(* IEC 61131-3 sources: daoli-st-library/DL_MathData (part 7) *)

(* ---- FC_DL_WaferCountYield.st ---- *)
(*==============================================================================
 * 组件名称 (Component)  : FC_DL_WaferCountYield
 * 所属子库 (Sublibrary) : DL_MathData
 * 当前版本 (Version)    : 1.0.0
 * 兼容性 (Platform)     : CODESYS 3.5 / TwinCAT 3 / 汇川 InoProShop / Machine Expert
 *                         仅依赖纯 IEC 61131-3 标准元素，零厂商方言
 * 功能描述 (Function)   : 晶圆投入/产出/返工三计数 → 良率百分数与损失分档。
 *                         良率 = 良品/投入 x 100；分档：A 级 >= 99、B 级 >= 95、
 *                         C 级 >= 90、D 级 < 90。纯函数无状态保持。
 * 溯源 (Origin)         : 道莅 clean-room 防御性实现
 * 本文件内含 (Contains) : TYPE E_DL_YieldGrade / TYPE E_DL_WaferErr /
 *                         FUNCTION FC_DL_WaferCountYield
 * 依赖 (Depends)        : 无 DL_ 内部依赖；仅 IEC 61131-3 标准元素
 * 红线自检 (Redline)    : 无外部全局变量、无硬件地址直引 ｜ 全变量中英双语同行注释
 *                         防除零 + 无符号减法先验下界防下溢 ｜ 枚举成员全部显式赋值
 *                         纯函数无状态保持 ｜ 输出在每条早退路径前已赋确定值
 * 错误码表 (Codes)      : 16#0001_0476 故障级(否) 成功
 *                         16#0001_0477 故障级 投入计数为 0（防除零拒绝）
 *                         16#0001_0478 故障级 良品计数大于投入计数（计数矛盾）
 *                         16#0001_0479 故障级 良品+返工大于投入（计数矛盾/下溢风险）
 *                         16#0001_047A 信息级 成功但落入 D 档（不置故障标志）
 * 修订历史 (Revision)   : 2026-11-17  v1.0.0  首版入库 · R27 · 阶段三批 1
 * 验收向量 (Acceptance) : input=1000, good=995, rework=3 → 良率 99.5% → A 档 0476
 *                         input=0 → 0477；good=1001>input=1000 → 0478；
 *                         good=990+rework=20>input=1000 → 0479；input=100,good=80 → D 档 047A
 *============================================================================*)

(*-----------------------------------------------------------------------------
 * 枚举: E_DL_YieldGrade（归属 DL_MathData，损失分档结果）
 *----------------------------------------------------------------------------*)
TYPE E_DL_YieldGrade :
(
    eGradeA := 0,    // A 档：良率 >= 99% / Grade A: yield at least 99 percent
    eGradeB := 1,    // B 档：良率 >= 95% 且 < 99% / Grade B: 95 to below 99 percent
    eGradeC := 2,    // C 档：良率 >= 90% 且 < 95% / Grade C: 90 to below 95 percent
    eGradeD := 3     // D 档：良率 < 90% / Grade D: below 90 percent
);
END_TYPE

(*-----------------------------------------------------------------------------
 * 枚举: E_DL_WaferErr（归属 DL_MathData，与 FC_DL_WaferCountYield 同文件）
 *----------------------------------------------------------------------------*)
TYPE E_DL_WaferErr :
(
    eOk           := 16#0001_0476,   // 成功 / Success
    eInputZero    := 16#0001_0477,   // 故障级：投入为 0，防除零拒绝 / Fault: zero input rejected
    eGoodOverIn   := 16#0001_0478,   // 故障级：良品大于投入 / Fault: good count exceeds input
    eCountContrad := 16#0001_0479,   // 故障级：良品+返工大于投入 / Fault: good plus rework exceeds input
    eGradeDNote   := 16#0001_047A    // 信息级：成功但 D 档 / Info: success but grade D
);
END_TYPE

(*==============================================================================
 * 函数: FC_DL_WaferCountYield（纯函数，无任何状态保持）
 * 调用约定: 每周期按需调用；bValid = 计数合法且结果可用。
 *============================================================================*)
FUNCTION FC_DL_WaferCountYield : BOOL
VAR_INPUT
    uInputCnt   : UDINT;               // 投入片数 [片]，有效域 0~1.0E9 / Wafer input count [pcs]
    uOutputGood : UDINT;               // 良品片数 [片] / Good wafer count [pcs]
    uReworkCnt  : UDINT;               // 返工片数 [片] / Rework wafer count [pcs]
END_VAR
VAR_OUTPUT
    fYieldPct   : REAL;                // 良率 [百分数] / Yield [percent]
    eGrade      : E_DL_YieldGrade;     // 损失分档 A~D / Yield grade A to D
    bValid      : BOOL;                // 输入合法且结果可用标志 / Input legal and result usable flag
    eError      : E_DL_WaferErr;       // 错误码 / Error code
END_VAR
VAR CONSTANT
    DL_WFR_INPUT_MAX  : UDINT := 1000000000;  // 投入计数上限 [片] / Input count upper bound [pcs]
    DL_WFR_GRADE_A    : REAL := 99.0;         // A 档门限 [百分数] / Grade A threshold [percent]
    DL_WFR_GRADE_B    : REAL := 95.0;         // B 档门限 [百分数] / Grade B threshold [percent]
    DL_WFR_GRADE_C    : REAL := 90.0;         // C 档门限 [百分数] / Grade C threshold [percent]
    DL_WFR_PCT        : REAL := 100.0;        // 百分数系数 [百分数] / Percent factor [percent]
    DL_WFR_ZERO       : REAL := 0.0;          // 零值常量，避免裸字面量 / Zero constant
END_VAR
VAR
    fYieldCalc : REAL;                 // 良率中间量 [百分数] / Yield intermediate [percent]
    uLossCnt   : UDINT;                // 损失片数 = 投入-良品-返工（校验后计算）[片] / Loss count [pcs]
END_VAR

(*------------------------------------------------------------------------------
 * 段 1｜出口默认值：任何早退路径前输出已确定（哨兵 0 良率 + D 档 + 无效）
 *----------------------------------------------------------------------------*)
FC_DL_WaferCountYield := FALSE;                     // 返回值默认无效 / return defaults to invalid
fYieldPct := DL_WFR_ZERO;                           // 良率哨兵 0（防除零语义：保持 0）/ yield sentinel zero
eGrade := E_DL_YieldGrade.eGradeD;                  // 分档哨兵 D 档 / grade sentinel D
bValid := FALSE;                                    // 合法标志默认 FALSE / validity defaults FALSE
eError := E_DL_WaferErr.eInputZero;                 // 默认投入为 0 码 / default zero-input code

(*------------------------------------------------------------------------------
 * 段 2｜投入为 0 闸：防除零拒绝（良率保持哨兵 0）
 *----------------------------------------------------------------------------*)
IF (uInputCnt = 0) OR (uInputCnt > DL_WFR_INPUT_MAX) THEN
    eError := E_DL_WaferErr.eInputZero;             // 故障级：投入为 0 或越上限 / fault: zero or out-of-range input
    RETURN;
END_IF

(*------------------------------------------------------------------------------
 * 段 3｜计数矛盾闸：良品不得大于投入；良品+返工不得大于投入（先验下界防下溢）
 *----------------------------------------------------------------------------*)
IF uOutputGood > uInputCnt THEN
    eError := E_DL_WaferErr.eGoodOverIn;            // 故障级：良品 > 投入 / fault: good exceeds input
    RETURN;
END_IF
IF uReworkCnt > (uInputCnt - uOutputGood) THEN      // 减法前已证 input >= good，无下溢 / no underflow, proven
    eError := E_DL_WaferErr.eCountContrad;          // 故障级：良品+返工 > 投入 / fault: count contradiction
    RETURN;
END_IF

(*------------------------------------------------------------------------------
 * 段 4｜良率计算与分档：fYield = good/input x 100（除子已证非零）
 *----------------------------------------------------------------------------*)
fYieldCalc := UDINT_TO_REAL(uOutputGood) / UDINT_TO_REAL(uInputCnt) * DL_WFR_PCT;   // 良率 [百分数] / yield [percent]
IF fYieldCalc > DL_WFR_PCT THEN
    fYieldCalc := DL_WFR_PCT;                       // 上限防护（计数矛盾已拦，兜底）/ ceiling guard
END_IF
fYieldPct := fYieldCalc;                            // 输出良率 / yield output
uLossCnt := uInputCnt - uOutputGood - uReworkCnt;   // 损失片数 [片]（两条矛盾闸已保证非负）/ loss count, proven non-negative
IF fYieldPct >= DL_WFR_GRADE_A THEN
    eGrade := E_DL_YieldGrade.eGradeA;              // A 档 / grade A
    eError := E_DL_WaferErr.eOk;                    // 成功码 / success code
ELSIF fYieldPct >= DL_WFR_GRADE_B THEN
    eGrade := E_DL_YieldGrade.eGradeB;              // B 档 / grade B
    eError := E_DL_WaferErr.eOk;                    // 成功码 / success code
ELSIF fYieldPct >= DL_WFR_GRADE_C THEN
    eGrade := E_DL_YieldGrade.eGradeC;              // C 档 / grade C
    eError := E_DL_WaferErr.eOk;                    // 成功码 / success code
ELSE
    eGrade := E_DL_YieldGrade.eGradeD;              // D 档 / grade D
    eError := E_DL_WaferErr.eGradeDNote;            // 信息级：成功但 D 档（损失片数佐证）/ info: grade D note
END_IF
bValid := TRUE;                                     // 输入合法，结果可用 / input legal, result usable
FC_DL_WaferCountYield := TRUE;                      // 返回有效 / return valid
RETURN;
END_FUNCTION

(* ---- FC_DL_AbsEx.st ---- *)
(*
    FC_DL_AbsEx —— 实数绝对值防御包装（-0.0 归一、NaN/无穷拦截、极值溢出钳位）
    ------------------------------------------------------------------
    分类      : DL_MathData / Math-Exp
    前缀      : FC_DL_
    版本      : 1.0.0
    溯源      : IEC 61131-3 标准语义的道莅防御性实现
                （内部委托平台内建函数，外围统一错误码/钳位/双语文档；
                  未复制任何闭源厂商源码，参考实现仅限 MIT/Apache 许可）
    平台      : 纯 IEC 61131-3，CODESYS / TwinCAT / InoProShop 通用
    作者      : 道莅代码库 · PLC编程专家（R15）
    ------------------------------------------------------------------
    功能说明  : 求输入实数的绝对值。NaN 输入直接拦截返回 0.0 并置 16#0001_015E；
                无穷输入（超出双精度有限极值）同口径拦截归零；-0.0 归一
                为 +0.0；负数经符号取反实现，当绝对值恰为双精度极值
                1.7976931348623157E308 时按上溢口径钳位到同值并置 16#0001_022C
                （钳位值与真实绝对值一致，bValid=TRUE 降级可用）。
                全程绝不向下游输出 NaN/Inf 毒值。
    错误码    : 0000 正常 / 16#0001_015E 入参越界（NaN/无穷，已归零） / 16#0001_022C 上溢下溢（已钳位到类型极值）
    修订记录  : 2026-11-16 v1.0.0 首次入库（R15）
*)
FUNCTION FC_DL_AbsEx : LREAL
VAR_INPUT
    lrIn : LREAL; // 输入实数 [无量纲]，任意有限值或 NaN/无穷 / input real value [dimensionless], any finite value or NaN/inf
END_VAR
VAR_OUTPUT
    eErr : UDINT; // 错误码，0=正常，1=入参越界，2=上溢钳位 / error id, 0=ok, 1=input out of domain, 2=overflow clamped
    bError   : BOOL; // 是否出错，eErr 非 0 时为 TRUE / error flag, TRUE when eErr is nonzero
    bValid   : BOOL; // 输出是否有效可用，16#0001_022C 钳位降级时保持 TRUE / output valid, stays TRUE for usable clamped result of code 2
END_VAR
VAR
    lrAbs : LREAL; // 绝对值中间量 [无量纲] / intermediate absolute value [dimensionless]
END_VAR
VAR CONSTANT
    DL_AB_MAXREAL : LREAL := 1.7976931348623157E308; // 双精度有限极值 [无量纲]，超界判无穷，禁魔法数 / double precision finite max [dimensionless], beyond treated as infinity, no magic numbers
END_VAR

// 段 1｜返回值与错误状态预置，任何早退路径不留脏码 / segment 1, preset return value and error states so no early exit leaves stale codes
FC_DL_AbsEx := 0.0; // 返回值预置安全值 0.0 [无量纲] / preset return to safe value 0.0
eErr    := 16#0000_0000; // 错误码预置正常 / preset error id to ok
bError      := FALSE; // 错误标志预置无错 / preset error flag to FALSE
bValid      := TRUE; // 有效标志预置可用 / preset valid flag to TRUE

// 段 2｜非有限拦截：NaN 用自不等判据，无穷用超极值判据，一律不进取反运算 / segment 2, non-finite interception, NaN by self-inequality and infinity by bound test
IF (lrIn <> lrIn) OR (lrIn > DL_AB_MAXREAL) OR (lrIn < -DL_AB_MAXREAL) THEN
    eErr := 16#0001_015E; // 信息级：输入非有限，已归零 / informational, non-finite input, zeroed
    bError   := TRUE; // 置错误标志 / raise error flag
    bValid   := FALSE; // 输出 0.0 非真实结果，不可用 / output 0.0 is not the true result, invalid
    RETURN; // 返回预置安全值 0.0 / return preset safe value 0.0
END_IF

// 段 3｜零值归一：与 0.0 精确比较对 -0.0 与 +0.0 均成立，统一归 +0.0 / segment 3, zero normalization, exact compare catches both minus zero and plus zero
IF lrIn = 0.0 THEN
    FC_DL_AbsEx := 0.0; // -0.0 归一为 +0.0 / normalize minus zero to plus zero
    RETURN;
END_IF

// 段 4｜负数取反与极值溢出钳位 / segment 4, negation for negative input with extreme-value overflow clamp
IF lrIn < 0.0 THEN
    IF lrIn <= -DL_AB_MAXREAL THEN
        lrAbs    := DL_AB_MAXREAL; // 绝对值恰为极值，按上溢口径钳位 / magnitude at the extreme, clamped per overflow policy
        eErr := 16#0001_022C; // 上溢码：已钳位到类型极值 / overflow code, clamped to type extreme
        bError   := TRUE; // 置错误标志 / raise error flag
        // bValid 保持 TRUE：钳位值与真实绝对值一致，降级可用 / valid stays TRUE, clamped value equals the true absolute value
    ELSE
        lrAbs := -lrIn; // 域内负数直接取反 / in-domain negative input negated
    END_IF
ELSE
    lrAbs := lrIn; // 正数直通 / positive input passes through
END_IF

// 段 5｜结果非有限复检兜底（防御纵深，正常路径不可达） / segment 5, result finiteness recheck as defense in depth
IF lrAbs <> lrAbs THEN
    lrAbs    := 0.0; // 兜底安全值 / bottom-line safe value
    eErr := 16#0001_015E; // 信息级：结果异常归零 / informational, abnormal result zeroed
    bError   := TRUE; // 置错误标志 / raise error flag
    bValid   := FALSE; // 输出不可用 / output invalid
END_IF
FC_DL_AbsEx := lrAbs; // 输出绝对值 [无量纲] / output the absolute value
END_FUNCTION

(* ---- FC_DL_AcosDegChk.st ---- *)
(*==============================================================================
 * 名称 : FC_DL_AcosDegChk —— 反余弦 → 角度（输入钳位 [-1,1]，越界仍按钳位计算）
 * 分类 / 前缀 / 版本 : DL_MathData / FC_DL_ / 1.0.0
 * 溯源 : 开源语义参考（OSCAT/AixOCAT 族，MIT）或 clean-room IEC 实现，未复制源码
 * 平台 : 纯 IEC 61131-3
 * 功能说明 : 返回 acos(x) 的角度制结果 [0,180]。输入越出 [-1,1] 时钳位到
 *            边界后仍按钳位值计算（bValid=FALSE、eErr 置码提示越界），不产生
 *            NaN。恒等式 acos(x)=atan2(sqrt(1-x^2), x)（弧度）转角度输出，
 *            纯 ATAN2/SQRT 内联实现，无库内跨件依赖。
 *            边界处理：输入非有限（NaN/±Inf）置 eErr 返回 0.0（不钳位计算）。
 * 错误码 : 16#0001_1B0D = 输入越出 [-1,1]（已钳位计算），或输入非有限（NaN/±Inf）
 *          eErr=0 且 bValid=TRUE 表示输入在域内、返回值可用
 * 状态机 : R6 标注 N/A（纯函数无顺序状态，以本节替代 ELSE 兜底）
 * 红线 : R1/R2/R3 ✓ 零全局/零IO/纯IEC ｜ R4 ✓ 非有限拦截/域钳位防 NaN ｜ R10 ✓ 标准转换 ｜ R11 ✓ 分号收尾 ｜ R15 ✓ 无保留字撞名
 * 修订记录 : 2026-11-23 v1.0.0 首次入库（R76）
 *============================================================================*)
FUNCTION FC_DL_AcosDegChk : LREAL
VAR_INPUT
    fX : LREAL;    // 余弦值输入 [-1,1]，越界钳位 / cosine value input, clamped into [-1,1]
END_VAR
VAR_OUTPUT
    eErr   : UDINT;    // 故障码，0=正常，1B0D=越界钳位或非有限 / error code
    bError : BOOL;     // TRUE=本件发生故障 / TRUE when fault occurred
    bValid : BOOL;     // TRUE=输入在域内且返回值可用 / TRUE when input in domain and result usable
END_VAR
VAR
    _x  : LREAL;       // 钳位后的输入 [无量纲] / clamped input
    _fR : LREAL;       // 弧度制反余弦结果 [rad] / arccosine result in radians
END_VAR

FC_DL_AcosDegChk := 0.0;                     // 返回值预设 0.0 / preset return to zero
eErr   := 16#0000_0000;                      // 故障码清零 / clear error code
bError := FALSE;                             // 故障标志清零 / clear error flag
bValid := TRUE;                              // 预设输出可用 / preset valid flag

IF (fX <> fX) OR ((fX - fX) <> (fX - fX)) THEN    // NaN 或 ±Inf / NaN or infinite
    eErr   := 16#0001_1B0D;                  // 置非有限故障码 / set non-finite code
    bError := TRUE;                          // 置故障标志 / set error flag
    bValid := FALSE;                         // 返回值不可用 / return not usable
    RETURN;                                  // 返回 0.0 / return zero
END_IF

_x := fX;                                    // 取输入 / take input
IF _x > 1.0 THEN                             // 上越界钳位 / clamp upper
    _x := 1.0;                               // 钳到 +1 / clamp to +1
    eErr   := 16#0001_1B0D;                  // 置越界码 / set out-of-domain code
    bError := TRUE;                          // 置故障标志 / set error flag
    bValid := FALSE;                         // 提示越界（仍按钳位值出结果）/ flag clamped compute
ELSIF _x < -1.0 THEN                         // 下越界钳位 / clamp lower
    _x := -1.0;                              // 钳到 -1 / clamp to -1
    eErr   := 16#0001_1B0D;                  // 置越界码 / set out-of-domain code
    bError := TRUE;                          // 置故障标志 / set error flag
    bValid := FALSE;                         // 提示越界（仍按钳位值出结果）/ flag clamped compute
END_IF

_fR := ATAN2(SQRT(1.0 - _x * _x), _x);       // acos(x)=atan2(sqrt(1-x^2),x)，弧度 / arccosine via atan2
FC_DL_AcosDegChk := _fR * 180.0 / 3.14159265358979323846;    // 弧度转角度 / radians to degrees

END_FUNCTION

(* ---- FC_DL_AcosEx.st ---- *)
(*
    FC_DL_AcosEx —— 反余弦防御包装（定义域 [-1,1] 域闸钳位 + NaN 拦截）
    ------------------------------------------------------------------
    分类      : DL_MathData / Math-Trig
    前缀      : FC_DL_
    版本      : 1.0.0
    溯源      : IEC 61131-3 标准语义的道莅防御性实现
                （内部委托平台内建函数，外围统一错误码/钳位/双语文档；
                  未复制任何闭源厂商源码，参考实现仅限 MIT/Apache 许可）
    平台      : 纯 IEC 61131-3，CODESYS / TwinCAT / InoProShop 通用
    作者      : 道莅代码库 · PLC编程专家（R15）
    ------------------------------------------------------------------
    功能说明  : 求输入的反余弦，返回值域 [0, pi]。与 FC_DL_AsinEx 同一
                钳位策略：NaN 输入拦截返回 0.0 并置 16#0001_0172；定义域 [-1,1]
                之外（含无穷）钳位到 ±1 并置 16#0001_0172，bValid=FALSE 但仍返回
                钳位后的计算结果（0 或 pi）供降级使用；入参为 0 时结果
                pi/2 属正常域内输出不置码；域内委托内建 ACOS，结果再做
                NaN 复检兜底。
    错误码    : 0000 正常 / 16#0001_0172 入参越界（NaN 已归零，或域外已钳位到 ±1）
    修订记录  : 2026-11-16 v1.0.0 首次入库（R15）
*)
FUNCTION FC_DL_AcosEx : LREAL
VAR_INPUT
    lrIn : LREAL; // 输入实数 [无量纲]，定义域 [-1,1] / input real value [dimensionless], domain minus 1 to plus 1
END_VAR
VAR_OUTPUT
    eErr : UDINT; // 错误码，0=正常，1=入参越界（已钳位/归零） / error id, 0=ok, 1=input out of domain, clamped or zeroed
    bError   : BOOL; // 是否出错，eErr 非 0 时为 TRUE / error flag, TRUE when eErr is nonzero
    bValid   : BOOL; // 输出是否有效可用，钳位/归零降级时为 FALSE / output valid, FALSE for clamped or zeroed degraded results
END_VAR
VAR
    lrUse : LREAL; // 钳位后的实际计算入参 [无量纲] / clamped value actually fed to the kernel [dimensionless]
END_VAR
VAR CONSTANT
    DL_AC_DOM : LREAL := 1.0; // 定义域边界 [无量纲]，闭区间 / domain bound [dimensionless], closed interval
END_VAR

// 段 1｜返回值与错误状态预置，任何早退路径不留脏码 / segment 1, preset return value and error states
FC_DL_AcosEx := 0.0; // 返回值预置安全值 0.0 / preset return to safe value 0.0
eErr    := 16#0000_0000; // 错误码预置正常 / preset error id to ok
bError      := FALSE; // 错误标志预置无错 / preset error flag to FALSE
bValid      := TRUE; // 有效标志预置可用 / preset valid flag to TRUE

// 段 2｜NaN 拦截：自不等判据，归零早退，不进内核 / segment 2, NaN interception by self-inequality, zeroed early exit
IF lrIn <> lrIn THEN
    eErr := 16#0001_0172; // 信息级：输入 NaN，已归零 / informational, NaN input, zeroed
    bError   := TRUE; // 置错误标志 / raise error flag
    bValid   := FALSE; // 输出不可用 / output invalid
    RETURN; // 返回预置安全值 0.0 / return preset safe value 0.0
END_IF

// 段 3｜定义域闸门：域外（含无穷）钳位到 ±1，仍返回钳位后结果 / segment 3, domain gate, out-of-domain including infinity clamped to plus or minus 1 with result still returned
IF lrIn > DL_AC_DOM THEN
    lrUse    := DL_AC_DOM; // 上越界钳位 +1 / upper overflow clamped to plus 1
    eErr := 16#0001_0172; // 信息级：域外已钳位 / informational, out of domain clamped
    bError   := TRUE; // 置错误标志 / raise error flag
    bValid   := FALSE; // 钳位结果非真实值 / clamped result is not the true value
ELSIF lrIn < -DL_AC_DOM THEN
    lrUse    := -DL_AC_DOM; // 下越界钳位 -1 / lower overflow clamped to minus 1
    eErr := 16#0001_0172; // 信息级：域外已钳位 / informational, out of domain clamped
    bError   := TRUE; // 置错误标志 / raise error flag
    bValid   := FALSE; // 钳位结果非真实值 / clamped result is not the true value
ELSE
    lrUse := lrIn; // 域内直通（0 输入得 pi/2 属正常） / in-domain pass-through, zero input yields pi over 2 normally
END_IF

// 段 4｜委托内建 ACOS / segment 4, delegation to built-in ACOS
FC_DL_AcosEx := ACOS(lrUse); // 委托内建 ACOS 内核 / delegate to built-in ACOS kernel

// 段 5｜结果 NaN 复检兜底（防御纵深，正常路径不可达） / segment 5, result NaN recheck as defense in depth
IF FC_DL_AcosEx <> FC_DL_AcosEx THEN
    FC_DL_AcosEx := 0.0; // 兜底安全值 / bottom-line safe value
    IF eErr = 16#0000_0000 THEN
        eErr := 16#0001_0172; // 首事件优先置码 / first-event priority code
        bError   := TRUE; // 置错误标志 / raise error flag
        bValid   := FALSE; // 输出不可用 / output invalid
    END_IF
END_IF
END_FUNCTION

(* ---- FC_DL_AcosSafe.st ---- *)
(*
    FC_DL_AcosSafe —— 反余弦 Safe 族防御包装（域钳位 + bClamped 显式标志 + 委托内建）
    ------------------------------------------------------------------
    分类      : DL_MathData / Math-Trig
    前缀      : FC_DL_
    版本      : 1.0.0
    来源标签  : iec-std-wrapper（T0）
    溯源      : IEC 61131-3 标准语义的道莅防御性实现
                （内部委托平台内建 ACOS，外围钳位/错误码/双语文档；
                  未复制任何闭源厂商源码）
    平台      : 纯 IEC 61131-3，CODESYS / TwinCAT / InoProShop 通用
    分工声明  : 与 FC_DL_AsinSafe 为镜像件（ACOS 口径），与存量 FC_DL_AcosEx
                分工——AcosEx 为码位族，本件为 Safe 族样板（bClamped 显式
                钳位标志 + 16#0002 子带码位）；边界验证向量取 ±1 两点。
    作者      : 道莅代码库 · PLC 编程专家（R57）
    ------------------------------------------------------------------
    功能说明  : 求输入的反余弦，返回值域 [0, pi]。四段式防御（R45）：
                NaN 双判据拦截归零早退；|x|>1（含无穷）钳到 ±1 并置 bClamped
                仍返回钳位结果供降级（边界向量 ±1 为合法输入直通）；
                域内委托内建 ACOS；结果 NaN 复检兜底。
    错误码    : 0000 正常 / 16#0002_0001 入参非有限已归零 / 16#0002_0002 域外已钳位
    修订记录  : 2026-11-21 v1.0.0 首次入库（R57 批 2 · 序号 7）
*)
FUNCTION FC_DL_AcosSafe : LREAL
VAR_INPUT
    lrIn : LREAL; // 输入实数 [无量纲]，定义域 [-1,1] / input real value [dimensionless], domain minus one to plus one
END_VAR
VAR_OUTPUT
    eErr     : UDINT; // 错误码，0 = 正常 / error code, zero is ok
    bError   : BOOL;  // 出错标志，eErr 非 0 时为真 / error flag, true when eErr is nonzero
    bValid   : BOOL;  // 结果是否为真实值，钳位/归零降级时为假 / the result is the true value, false when degraded
    bClamped : BOOL;  // 本次调用发生定义域钳位 [-] / a domain clamp happened this call
END_VAR
VAR
    lrUse : LREAL; // 钳位后的实际计算入参 [无量纲] / the clamped value fed to the kernel [dimensionless]
END_VAR
VAR CONSTANT
    DL_ACS_DOM : LREAL := 1.0; // 定义域边界 [无量纲]，闭区间 / the domain bound [dimensionless], closed interval
END_VAR

// 段 1｜返回值与错误状态预置安全值（四段式第一段，R45）/ segment 1, preset the return and error states
FC_DL_AcosSafe := 0.0; // 返回值预置安全值 0.0 / preset the return to the safe zero
eErr     := 16#0000_0000; // 错误码预置正常 / preset the code to ok
bError   := FALSE; // 错误标志预置假 / preset the error flag false
bValid   := TRUE; // 有效标志预置真 / preset the valid flag true
bClamped := FALSE; // 钳位标志预置假 / preset the clamp flag false

// 段 2｜非有限拦截（双判据）：命中不调内建直接早退 / segment 2, the non finite interception
IF (lrIn <> lrIn) OR ((lrIn - lrIn) <> (lrIn - lrIn)) THEN // NaN 或无穷 / NaN or infinity
    eErr   := 16#0002_0001; // 信息级：输入非有限已归零 / informational, a non finite input zeroed
    bError := TRUE; // 置错误标志 / raise the error flag
    bValid := FALSE; // 输出不可用 / the output void
    RETURN; // 返回预置安全值 0.0 / return the preset safe zero
END_IF

// 段 3｜定义域闸门：域外钳到 ±1 并置 bClamped（±1 两边界点为合法输入直通）/ segment 3, the domain gate, the boundary points plus or minus one legal
IF lrIn > DL_ACS_DOM THEN // 上越界 / above the bound
    lrUse    := DL_ACS_DOM; // 钳到 +1 / clamp to plus one
    eErr     := 16#0002_0002; // 信息级：域外已钳位 / informational, clamped
    bError   := TRUE; // 置错误标志 / raise the error flag
    bValid   := FALSE; // 钳位结果非真实值 / the clamped result is not the true value
    bClamped := TRUE; // 置钳位标志 / raise the clamp flag
ELSIF lrIn < -DL_ACS_DOM THEN // 下越界 / below the bound
    lrUse    := -DL_ACS_DOM; // 钳到 -1 / clamp to minus one
    eErr     := 16#0002_0002; // 信息级：域外已钳位 / informational, clamped
    bError   := TRUE; // 置错误标志 / raise the error flag
    bValid   := FALSE; // 钳位结果非真实值 / the clamped result is not the true value
    bClamped := TRUE; // 置钳位标志 / raise the clamp flag
ELSE // 域内直通 / inside the domain
    lrUse := lrIn; // 直通 / passthrough
END_IF

// 段 4｜委托内建 ACOS（禁重实现数学内核）/ segment 4, delegation to the built-in ACOS
FC_DL_AcosSafe := ACOS(lrUse); // 委托内建内核 / delegate to the built-in kernel

// 段 5｜结果 NaN 复检兜底（防御纵深，正常路径不可达）/ segment 5, the result recheck as defense in depth
IF (FC_DL_AcosSafe <> FC_DL_AcosSafe) OR ((FC_DL_AcosSafe - FC_DL_AcosSafe) <> (FC_DL_AcosSafe - FC_DL_AcosSafe)) THEN // 结果非有限 / a non finite result
    FC_DL_AcosSafe := 0.0; // 兜底安全值 / the bottom-line safe value
    IF eErr = 16#0000_0000 THEN // 首事件优先置码 / the first event keeps the code
        eErr   := 16#0002_0001; // 信息级：结果非有限已归零 / informational, a non finite result zeroed
        bError := TRUE; // 置错误标志 / raise the error flag
        bValid := FALSE; // 输出不可用 / the output void
    END_IF
END_IF
END_FUNCTION

(* ---- FC_DL_Affine2Apply.st ---- *)
//==============================================================================
// 函数：FC_DL_Affine2Apply ｜ 中文名称：二维仿射矩阵对点坐标应用
// 所属子库：DL_MathData ｜ 版本：v1.0.0 ｜ 兼容：CODESYS V3.5+ / TwinCAT 3 / 汇川 InoProShop
// 功能描述：单片 3x3 仿射矩阵对单点坐标 (x, y) 应用变换，p' = M x [x, y, 1]^T
//           （列向量右乘，与 FC_DL_Affine2DCompose 的合成约定构成定义-应用
//           逆对：Compose 产出矩阵、Apply 消费矩阵）。现场语义：视觉像素
//           坐标到机械毫米坐标的单点映射、纠偏平台坐标换算、印刷套准偏移。
//           第三行偏差提示为本件信息级职责：喂入矩阵第三行偏离 (0, 0, 1)
//           超容差时按仿射截断（只用前两行），输出照算并提示，便于标定
//           链上游把透视矩阵误接进仿射链时尽早暴露。
// 开源溯源 (Origin)：道莅 clean-room 防御性实现（仅借 LGF 分类事实/参数域/行为定义，零代码行与符号名复制）
// 单位表：点坐标[用户单位] / 矩阵线性块[无量纲] / 平移列[用户单位]
// 错误码表：16#0001_0469 信息级（矩阵第三行偏离 (0,0,1) 超容差，按仿射截断
//           照算，不置 bError）/ 16#0001_046A 预留禁用（不得挪用）/
//           16#0001_046B 预留禁用（不得挪用）/ 16#0001_03B9 故障级（任一
//           输入非有限，或结果非有限溢出，置 bError，输出 0）/
//           16#0001_03BA 预留禁用（不得挪用）
// 状态机：N/A——纯函数无顺序状态机，无 CASE 可写，非法状态不可能出现，以头注释说明替代 ELSE 兜底
// 边界行为：① 矩阵元素或点坐标非有限（NaN 自反判 + 幅值上限兜底，R79）→
//           故障 03B9、输出 0、bValid := FALSE；② 结果非有限（大坐标乘
//           大缩放溢出）→ 复用 03B9（R90：与输入非法共用「数据不可信」
//           语义，现有输出组合不可观测出独立信息，不新占码位）；
//           ③ 第三行偏差仅提示不阻断（信息 0469），仿射截断照算；
//           ④ 失能清零不适用（纯函数无使能闸，非法输入即故障早退）；
//           ⑤ 安全侧 = 故障路径输出 0 而非原坐标，禁止未变换坐标冒充
//           已变换坐标进入下游；
//           ⑥ 恒等矩阵输入时输出等于输入（数值恒等由乘 1.0 保证，
//           非位拷贝）。
// 验收向量（算法已证，手算）：① 恒等矩阵 + (3,4) → (3,4)；② 平移
//           (10,20) + (1,1) → (11,21)；③ 旋转 90 度 + (1,0) → (0,1)。
//           编译器已证（三平台）：未跑，由收口方登记。
// 修订历史：v1.0.0 2026-11-17 首版（R24 派单 · T2-1 LGF Math 仿射变换族）
//==============================================================================

FUNCTION FC_DL_Affine2Apply : BOOL
VAR_INPUT
    afM : ARRAY[0..2, 0..2] OF LREAL;       // 仿射变换矩阵 [无量纲+用户单位混合]，行主序，p' = M x p / Affine transform matrix, row-major
    fX  : LREAL;                            // 源点 X [用户单位] / Source point X [user unit]
    fY  : LREAL;                            // 源点 Y [用户单位] / Source point Y [user unit]
END_VAR
VAR_OUTPUT
    fOutX  : LREAL;                         // 变换后 X [用户单位] / Transformed X [user unit]
    fOutY  : LREAL;                         // 变换后 Y [用户单位] / Transformed Y [user unit]
    eErr   : UDINT;                         // 错误码，0 = 无错，码位 16#0001_0469 起信息级、16#0001_03B9 起故障级（分带见错误码表） / Error code, 0 = no error, band info/fault per the code table
    bError : BOOL;                          // 故障级标志，仅故障级错误置位 / Fault-class flag, set only on fault-level codes
    bValid : BOOL;                          // 结果可用标志 / Result usable flag
END_VAR
VAR CONSTANT
    DL_A2A_EPS      : LREAL := 1.0E-6;      // 第三行偏差容差与浮点判零共用 [无量纲] / Third-row deviation and zero tolerance [dimensionless]
    DL_A2A_INF      : LREAL := 1.7976931348623157E308; // LREAL 幅值上限 / LREAL magnitude ceiling
    DL_A2A_ZERO     : LREAL := 0.0;         // 零值常量，避免裸字面量 [无量纲] / Zero constant, avoids a bare literal [dimensionless]
    DL_A2A_ONE      : LREAL := 1.0;         // 单位常量，第三行齐次项期望值 [无量纲] / Unity constant, expected homogeneous entry [dimensionless]
END_VAR
VAR
    fXt     : LREAL;                        // 第一行点积暂存 [用户单位] / First-row dot product staging
    fYt     : LREAL;                        // 第二行点积暂存 [用户单位] / Second-row dot product staging
    bNonFin : BOOL;                         // 非有限判定中间标志 / Non-finite detection intermediate flag
    nI      : INT;                          // 行循环索引 [—] / Row loop index
    nJ      : INT;                          // 列循环索引 [—] / Column loop index
END_VAR

(*------------------------------------------------------------------------------
 * 段 1｜出口默认值：返回值与输出预置（安全侧 = 0）
 *      Exit defaults: return value and outputs preset, fail-safe zero
 *-----------------------------------------------------------------------------*)
FC_DL_Affine2Apply := FALSE;                // 返回值默认无效 / Return value preset invalid
fOutX := DL_A2A_ZERO;                       // 输出 X 预置 0 / Preset X to zero
fOutY := DL_A2A_ZERO;                       // 输出 Y 预置 0 / Preset Y to zero
eErr   := 16#0000_0000;                     // 错误码先清零 / Error code cleared first
bError := FALSE;                            // 故障标志先清零 / Fault flag cleared first
bValid := FALSE;                            // 可用标志先清零 / Usable flag cleared first

(*------------------------------------------------------------------------------
 * 段 2｜输入非有限闸：矩阵九元素 + 点坐标（R79 双侧幅值判）
 *      Input non-finite gate over nine matrix entries and the point
 *-----------------------------------------------------------------------------*)
bNonFin := (fX <> fX) OR (ABS(fX) > DL_A2A_INF)
        OR (fY <> fY) OR (ABS(fY) > DL_A2A_INF); // 点坐标非有限判定 / Point non-finite check
FOR nI := 0 TO 2 DO
    FOR nJ := 0 TO 2 DO
        IF (afM[nI, nJ] <> afM[nI, nJ]) OR (ABS(afM[nI, nJ]) > DL_A2A_INF) THEN
            bNonFin := TRUE;                // 命中非有限矩阵元素 / Non-finite matrix entry hit
        END_IF
    END_FOR
END_FOR
IF bNonFin THEN
    eErr   := 16#0001_03B9;                 // 故障级：输入非有限 / Fault: non-finite input
    bError := TRUE;                         // 置故障标志（R45 配对） / Raise the fault flag
    bValid := FALSE;                        // 输出不可用 / Outputs unusable
    RETURN;                                 // 故障早退，输出保持 0 / Early return, outputs stay zero
END_IF

(*------------------------------------------------------------------------------
 * 段 3｜仿射应用：只用前两行点积（第三行截断，见段 4 提示）
 *      Affine application, first two rows only
 *-----------------------------------------------------------------------------*)
fXt := afM[0, 0] * fX + afM[0, 1] * fY + afM[0, 2]; // 第一行点积 [用户单位] / First-row dot product
fYt := afM[1, 0] * fX + afM[1, 1] * fY + afM[1, 2]; // 第二行点积 [用户单位] / Second-row dot product

(*------------------------------------------------------------------------------
 * 段 4｜第三行偏差提示：偏离 (0, 0, 1) 超容差 → 信息 0469（照算不阻断）
 *      Third-row deviation notice, computation continues
 *-----------------------------------------------------------------------------*)
IF (ABS(afM[2, 0]) > DL_A2A_EPS) OR (ABS(afM[2, 1]) > DL_A2A_EPS)
   OR (ABS(afM[2, 2] - DL_A2A_ONE) > DL_A2A_EPS) THEN
    eErr := 16#0001_0469;                   // 信息级：第三行非标准仿射，已按仿射截断 / Info: non-standard third row, affine-truncated
END_IF

(*------------------------------------------------------------------------------
 * 段 5｜结果非有限复检：大缩放乘大坐标可能溢出（复用 03B9，R90）
 *      Result non-finite recheck, code reused per R90
 *-----------------------------------------------------------------------------*)
IF (fXt <> fXt) OR (ABS(fXt) > DL_A2A_INF)
   OR (fYt <> fYt) OR (ABS(fYt) > DL_A2A_INF) THEN
    fOutX := DL_A2A_ZERO;                   // 溢出即输出 0（安全侧） / Overflow yields zero
    fOutY := DL_A2A_ZERO;                   // 溢出即输出 0 / Overflow yields zero
    eErr   := 16#0001_03B9;                 // 故障级：结果溢出复用输入非法码（R90） / Fault: overflow, code reused per R90
    bError := TRUE;                         // 置故障标志 / Raise the fault flag
    bValid := FALSE;                        // 输出不可用 / Outputs unusable
    RETURN;                                 // 故障早退 / Early return
END_IF

(*------------------------------------------------------------------------------
 * 段 6｜出口
 *      Exit
 *-----------------------------------------------------------------------------*)
fOutX := fXt;                               // 变换后 X 出口 / Transformed X outlet
fOutY := fYt;                               // 变换后 Y 出口 / Transformed Y outlet
bValid := TRUE;                             // 结果可用（含 0469 提示情形） / Result usable, including the 0469 notice case
FC_DL_Affine2Apply := TRUE;                 // 返回 TRUE = 应用有效 / Return TRUE = application valid
END_FUNCTION

(* ---- FC_DL_Affine2DChain.st ---- *)
(*
  ==================================================================
  组件名 Component  : FC_DL_Affine2DChain
  分类   Category   : DL_MathData
  复杂度 Complexity  : 中
  版本   Version    : 1.0.1
  功能   Purpose    : N 级 2D 仿射链一次合成。输入 nCount 个 3×3 齐次矩阵，按
                      固定次序合成 MOut = Mn × … × M2 × M1（列向量约定，先施加
                      M1），中间任一奇异即整体失效并置故障码，不外泄半结果。
  来源   Source     : t2-1-lgf-math（LGF Math 仿射族多级链合成）
  溯源   Origin     : 矩阵链式合成属公开线性代数语义，clean-room 自研实现（逐级
                      委托本库 FC_DL_Affine2DCompose 内核），未复制任何厂商源码。
  平台   Platform   : 纯 IEC 61131-3（仅 FOR / 数组 / 委托调用），三平台通用
  分工声明 Split     : 与 FC_DL_Affine2DCompose（两级属主）互补——后者只合成
                      两级并负责行列式相对判据；本件做 N 级链调度、退化分支与
                      链级码位装配，不重实现乘法内核、不重声明任何矩阵类型。
  依赖     Depends  : FC_DL_Affine2DCompose（DL_MathData 属主，本件逐级委托）
  作者   Author     : 道莅代码库 · PLC 编程专家（R60）
  ------------------------------------------------------------------
  边界 Boundary     :
                      一 合成次序写死列向量约定 MOut = Mn × … × M1：M1 先施加，
                         Mn 后施加；调用方若要行向量约定须自行转置，本件不设开关；
                      二 链长退化显式：nCount ≤ 0 输出单位阵并置信息级码；nCount
                         超 8 级钳位续算并置信息级码（不静默截断）；
                      三 有限性闸逐个枚举浮点输入：本件声明区 LREAL 输入集合 =
                         afMats 的 9 × nCount 个元素，闸内逐元素引用同一集合，
                         无标量 LREAL 引脚（R272 覆盖自证：9×nUsed 全枚举）；
                      四 中途奇异或中途非有限即整体失效：bValid = FALSE、输出
                         保持单位阵（不外泄半结果），故障码一次锁存于本次调用；
                      五 只读输入矩阵，不改调用方数组（PercentileLReal 纪律）。
  错误码   Codes    :
    16#0001_0620【故障级】中间阵奇异或委托内核判不可用，链合成终止
    16#0001_0621【故障级】输入矩阵含非有限元素（NaN / Inf），链合成终止
    16#0001_0622【信息级】链长越域已钳位（≤0 出单位阵，>8 钳到 8 级）
  验收   Acceptance :
    算法已证（脚本）：未跑 ｜ 编译器已证（三平台）：未跑
    V1 两级：M1 平移 (1,2)、M2 缩放 ×2 → 单位点 (0,0) 过链得 (2,4)
    V2 nCount=0 → 单位阵、bValid=TRUE、码 0622
    V3 第二级首行全零（奇异）→ bValid=FALSE、码 0620、输出仍为单位阵
  修订记录 Revision  :
    2026-11-21  v1.0.0  R60 首版（批 2 · 序号 6）
    2026-11-21  v1.0.1  R61 返修：D5 累加器改单位阵起步、逐级全委托（含
                        nUsed=1 单级链奇异判，R284）；D6 信息级 0622 两处
                        不再置 bError（R285 口径统一）
  ==================================================================
*)
FUNCTION FC_DL_Affine2DChain : BOOL
VAR_IN_OUT
    afMats : ARRAY[0..7, 0..2, 0..2] OF LREAL; // 链矩阵组 [无量纲 + 用户单位混合]，行主序，第 0 级先施加 / the chain matrices, row major, level zero applied first
END_VAR
VAR_INPUT
    nCount : DINT; // 链级数 [级]，合法域 1..8 / the chain level count, legal from one to eight
END_VAR
VAR_OUTPUT
    afMOut : ARRAY[0..2, 0..2] OF LREAL; // 合成矩阵 [无量纲 + 用户单位混合] / the composed matrix
    bValid : BOOL;                       // 结果可用标志（链中任一级失效即假）[-] / the result usable flag
    eErr   : UDINT;                      // 错误码，0 = 正常 / the error code, zero is ok
    bError : BOOL;                       // 故障锁存标志 [-] / the fault flag
END_VAR
VAR
    afAcc     : ARRAY[0..2, 0..2] OF LREAL; // 累加矩阵（当前已合成结果） / the accumulator of the composed so far
    afTmp     : ARRAY[0..2, 0..2] OF LREAL; // 本级乘积暂存（检过才接替累加器） / the staging product of this level
    afMk      : ARRAY[0..2, 0..2] OF LREAL; // 本级矩阵切片副本（三维数组不可直接切片传参） / the slice copy of this level
    nLevel    : DINT;  // 级遍历索引 [级] / the level loop index
    nI        : DINT;  // 行索引 [行] / the row index
    nJ        : DINT;  // 列索引 [列] / the column index
    nUsed     : DINT;  // 钳位后的实际级数 [级] / the clamped level count
    bAbort    : BOOL;  // 链终止标志（有限闸或奇异闸命中）[-] / the chain abort flag
    bClamped  : BOOL;  // 链长钳位标记 [-] / the level clamp flag
    bSubValid : BOOL;  // 委托内核结果可用位 [-] / the delegate usable bit
    bSubErr   : BOOL;  // 委托内核故障位 [-] / the delegate fault bit
    uSubErr   : UDINT; // 委托内核错误码 [码] / the delegate error code
END_VAR
VAR CONSTANT
    DL_A2CH_CHMAX : DINT := 8; // 链级数上界 [级]，与数组第 1 维一致 / the level bound aligned with the first dimension
END_VAR

// 段 1｜返回值与错误状态预置安全值（四段式第一段，R45）+ 输出预置单位阵 / segment 1, the preset of the return, the codes and the identity matrix
FC_DL_Affine2DChain := FALSE; // 返回值预置假 / preset the return false
bValid := FALSE; // 有效标志预置假 / preset the validity false
eErr := 16#0000_0000; // 错误码预置正常 / preset the code to ok
bError := FALSE; // 故障标志预置假 / preset the error flag false
bAbort := FALSE; // 终止标志预置假 / preset the abort flag false
bClamped := FALSE; // 钳位标记预置假 / preset the clamp flag false
bSubValid := FALSE; // 委托有效位预置假 / preset the delegate usable bit false
bSubErr := FALSE; // 委托故障位预置假 / preset the delegate fault bit false
uSubErr := 16#0000_0000; // 委托码预置零 / preset the delegate code zero
nUsed := 0; // 实际级数预置零 / preset the used level zero
FOR nI := 0 TO 2 DO // 单位阵装配 / build the identity matrix
    FOR nJ := 0 TO 2 DO // 列遍历 / the column loop
        IF nI = nJ THEN // 主对角 / the main diagonal
            afMOut[nI, nJ] := 1.0; // 对角置一 / unit on the diagonal
            afAcc[nI, nJ] := 1.0; // 累加器同步置一 / the accumulator seeded the same
        ELSE // 非对角 / the off diagonal
            afMOut[nI, nJ] := 0.0; // 非对角置零 / zero off the diagonal
            afAcc[nI, nJ] := 0.0; // 累加器同步置零 / the accumulator seeded the same
        END_IF
        afTmp[nI, nJ] := 0.0; // 暂存阵清零 / clear the staging matrix
        afMk[nI, nJ] := 0.0; // 切片副本清零 / clear the slice copy
    END_FOR
END_FOR

// 段 2｜链长域闸（退化与钳位显式，边界二）/ segment 2, the level count gate with the explicit degenerate branch
IF nCount < 1 THEN // 链长为零或负：退化为单位阵 / a non positive count degenerates to the identity
    eErr := 16#0001_0622; // 信息级：链长越域已钳位（信息级不置 bError，R285 口径统一，D6 返修）/ informational, the level count clamped, no fault bit
    bValid := TRUE; // 单位阵是合法结果 / the identity is a legal result
    FC_DL_Affine2DChain := TRUE; // 返回成功 / return success
    RETURN; // 早退：afMOut 已为单位阵（段 1 预置）/ early return with the identity already preset
END_IF
nUsed := nCount; // 域内接管级数 / take the count inside the domain
IF nUsed > DL_A2CH_CHMAX THEN // 超上界 / above the bound
    nUsed := DL_A2CH_CHMAX; // 钳到 8 级 / clamp to eight levels
    bClamped := TRUE; // 置钳位标记 / raise the clamp flag
END_IF

// 段 3｜有限性闸：9 × nUsed 个浮点元素逐个枚举（R272 覆盖自证，边界三）/ segment 3, the finiteness gate over every enumerated element
FOR nLevel := 0 TO nUsed - 1 DO // 级遍历 / the level loop
    FOR nI := 0 TO 2 DO // 行遍历 / the row loop
        FOR nJ := 0 TO 2 DO // 列遍历 / the column loop
            IF (afMats[nLevel, nI, nJ] <> afMats[nLevel, nI, nJ])
            OR ((afMats[nLevel, nI, nJ] - afMats[nLevel, nI, nJ]) <> (afMats[nLevel, nI, nJ] - afMats[nLevel, nI, nJ])) THEN // NaN 自反判 + Inf 差值自减判 / the NaN reflexive and the Inf difference tests
                bAbort := TRUE; // 置终止标志 / raise the abort flag
            END_IF
        END_FOR
    END_FOR
END_FOR
IF bAbort THEN // 输入含非有限 / a non finite input exists
    eErr := 16#0001_0621; // 故障级：输入矩阵含非有限元素 / fault grade, a non finite element in the input
    bError := TRUE; // 置错误标志（R45 配对）/ raise the error flag, paired with the fault code
    bValid := FALSE; // 结果不可用 / the result void
    RETURN; // 早退：afMOut 保持单位阵（不外泄半结果，边界四）/ early return with the identity kept
END_IF

// 段 4｜逐级合成：MOut = Mn × … × M1（累加器以单位阵起步、逐级全委托；D5 返修：nUsed=1 单级链也走一次委托补奇异判，R284）/ segment 4, the per level composition, the accumulator starts from the identity and every level is delegated
FOR nLevel := 0 TO nUsed - 1 DO // 第 0..nUsed-1 级逐级合成（单位阵为左乘起点）/ compose from level zero with the identity seeded accumulator
  IF NOT bAbort THEN // 链未终止才继续合成（终止后不再用半结果继续乘）/ compose only while the chain is alive
    afMk[0, 0] := afMats[nLevel, 0, 0]; // 切片副本第 0 行第 0 列 / slice row zero column zero
    afMk[0, 1] := afMats[nLevel, 0, 1]; // 切片副本第 0 行第 1 列 / slice row zero column one
    afMk[0, 2] := afMats[nLevel, 0, 2]; // 切片副本第 0 行第 2 列 / slice row zero column two
    afMk[1, 0] := afMats[nLevel, 1, 0]; // 切片副本第 1 行第 0 列 / slice row one column zero
    afMk[1, 1] := afMats[nLevel, 1, 1]; // 切片副本第 1 行第 1 列 / slice row one column one
    afMk[1, 2] := afMats[nLevel, 1, 2]; // 切片副本第 1 行第 2 列 / slice row one column two
    afMk[2, 0] := afMats[nLevel, 2, 0]; // 切片副本第 2 行第 0 列 / slice row two column zero
    afMk[2, 1] := afMats[nLevel, 2, 1]; // 切片副本第 2 行第 1 列 / slice row two column one
    afMk[2, 2] := afMats[nLevel, 2, 2]; // 切片副本第 2 行第 2 列 / slice row two column two
    IF NOT FC_DL_Affine2DCompose(afM1 := afAcc, afM2 := afMk, afMOut => afTmp, eErr => uSubErr, bError => bSubErr, bValid => bSubValid) THEN // 委托两级内核（含行列式相对判据；nUsed=1 时 afAcc 为单位阵，单位阵左乘精确无损，单级奇异判由本次委托补齐，D5）/ delegate the two level kernel, the identity left multiply is exact
        bAbort := TRUE; // 本级不可用 / this level is unusable
    END_IF
    IF bAbort OR (NOT bSubValid) THEN // 奇异或不可用即整体终止 / a singular or unusable level aborts the chain
        bAbort := TRUE; // 锁住终止标志 / hold the abort flag
    ELSE // 本级通过：接替累加器 / this level passed, take over the accumulator
        afAcc[0, 0] := afTmp[0, 0]; // 累加器接替第 0 行第 0 列 / take over row zero column zero
        afAcc[0, 1] := afTmp[0, 1]; // 累加器接替第 0 行第 1 列 / take over row zero column one
        afAcc[0, 2] := afTmp[0, 2]; // 累加器接替第 0 行第 2 列 / take over row zero column two
        afAcc[1, 0] := afTmp[1, 0]; // 累加器接替第 1 行第 0 列 / take over row one column zero
        afAcc[1, 1] := afTmp[1, 1]; // 累加器接替第 1 行第 1 列 / take over row one column one
        afAcc[1, 2] := afTmp[1, 2]; // 累加器接替第 1 行第 2 列 / take over row one column two
        afAcc[2, 0] := afTmp[2, 0]; // 累加器接替第 2 行第 0 列 / take over row two column zero
        afAcc[2, 1] := afTmp[2, 1]; // 累加器接替第 2 行第 1 列 / take over row two column one
        afAcc[2, 2] := afTmp[2, 2]; // 累加器接替第 2 行第 2 列 / take over row two column two
    END_IF
  END_IF
END_FOR

// 段 5｜出口装配：仅在全链通过时外泄合成阵（边界四）/ segment 5, the outlet assembly, exported only when the whole chain passed
IF bAbort THEN // 链终止 / the chain aborted
    eErr := 16#0001_0620; // 故障级：中间阵奇异或不可用 / fault grade, a singular or unusable intermediate
    bError := TRUE; // 置错误标志（R45 配对）/ raise the error flag, paired with the fault code
    bValid := FALSE; // 结果不可用 / the result void
    FC_DL_Affine2DChain := FALSE; // 返回失败（afMOut 保持单位阵）/ return failure with the identity kept
ELSE // 全链通过 / the whole chain passed
    afMOut[0, 0] := afAcc[0, 0]; // 出口第 0 行第 0 列 / outlet row zero column zero
    afMOut[0, 1] := afAcc[0, 1]; // 出口第 0 行第 1 列 / outlet row zero column one
    afMOut[0, 2] := afAcc[0, 2]; // 出口第 0 行第 2 列 / outlet row zero column two
    afMOut[1, 0] := afAcc[1, 0]; // 出口第 1 行第 0 列 / outlet row one column zero
    afMOut[1, 1] := afAcc[1, 1]; // 出口第 1 行第 1 列 / outlet row one column one
    afMOut[1, 2] := afAcc[1, 2]; // 出口第 1 行第 2 列 / outlet row one column two
    afMOut[2, 0] := afAcc[2, 0]; // 出口第 2 行第 0 列 / outlet row two column zero
    afMOut[2, 1] := afAcc[2, 1]; // 出口第 2 行第 1 列 / outlet row two column one
    afMOut[2, 2] := afAcc[2, 2]; // 出口第 2 行第 2 列 / outlet row two column two
    bValid := TRUE; // 结果可用 / the result is usable
    FC_DL_Affine2DChain := TRUE; // 返回成功 / return success
    IF bClamped THEN // 链长被钳位 / the level count was clamped
        eErr := 16#0001_0622; // 信息级：链长越域已钳位（信息级不置 bError，R285 口径统一，D6 返修）/ informational, the level count clamped, no fault bit
    END_IF
END_IF
END_FUNCTION

(* ---- FC_DL_Affine2DCompose.st ---- *)
//==============================================================================
// 函数：FC_DL_Affine2DCompose ｜ 中文名称：二维仿射变换矩阵合成
// 所属子库：DL_MathData ｜ 版本：v1.0.0 ｜ 兼容：CODESYS V3.5+ / TwinCAT 3 / 汇川 InoProShop
// 功能描述：两片 3x3 仿射矩阵按「先施加 M1、后施加 M2」的次序合成为单片
//           矩阵 MOut = M2 x M1（本库点变换约定 p' = M x p，列向量右乘），
//           单次调用内完成 3x3 乘法、行列式可逆性校验与双向非有限复检。
//           现场语义：视觉标定链的多级坐标映射（像素→机械→工件）合并为
//           单矩阵、纠偏平台级联、平移/旋转/缩放/剪切的按序合成。
//           合成次序与列向量约定为本库自有规格；行列式 |det| 小于容差判
//           不可逆，按信息级降级输出（合成结果本身仍有效，仅其逆变换
//           不可用），故障级只留给非法输入与结果溢出。
//           第三行按仿射约定忽略（不校验 0/0/1），第三行偏差提示职责
//           归 FC_DL_Affine2Apply 承担，本件不重复占用码位（R90）。
// 开源溯源 (Origin)：道莅 clean-room 防御性实现（仅借 LGF 分类事实/参数域/行为定义，零代码行与符号名复制）
// 单位表：矩阵线性块元素[无量纲]（旋转/缩放/剪切）/ 平移列元素[用户单位]
// 错误码表：16#0001_0466 信息级（合成矩阵行列式 |det| < 容差，变换不可逆，
//           结果照常输出，不置 bError）/ 16#0001_0467 预留禁用（不得挪用）/
//           16#0001_0468 预留禁用（不得挪用）/ 16#0001_03B7 故障级（任一
//           输入矩阵元素非有限，或乘积结果非有限溢出，置 bError，输出
//           零矩阵）/ 16#0001_03B8 预留禁用（不得挪用）
// 状态机：N/A——纯函数无顺序状态机，无 CASE 可写，非法状态不可能出现，以头注释说明替代 ELSE 兜底
// 边界行为：① 任一输入元素非有限（NaN 用自反判 x <> x，Inf 用幅值上限
//           兜底，R79）→ 故障 03B7、输出零矩阵、bValid := FALSE；
//           ② 乘积结果非有限（大坐标乘大缩放溢出）→ 复用 03B7（R90：
//           该场景与输入非法共用「矩阵数据不可信」语义，现有输出组合
//           不可观测出独立信息，不新占码位）、输出零矩阵；
//           ③ 行列式绝对值 < 1E-6 → 信息 0466，结果照常输出（降级
//           可观测，不置 bError）；
//           ④ 失能清零不适用（纯函数无使能闸，非法输入即故障早退）；
//           ⑤ 安全侧 = 故障路径输出零矩阵而非原矩阵，禁止半合成残阵
//           外泄到下游点应用件；
//           ⑥ 第三行不参与合成合法性判定：乘法仍按完整 3x3 执行，第三
//           行结果照算输出，调用方若喂入非标准第三行由 Apply 侧提示。
// 验收向量（算法已证，手算）：① M1=绕原点旋转 90 度、M2=平移 (10,0) →
//           MOut 平移列 = (0,10)、线性块为旋转 90 度；② M1=M2=恒等 →
//           MOut=恒等；③ M1 含缩放 (2,0.5)、M2 含剪切 k=1 → det(MOut)
//           = 2x0.5 = 1（合成保序：det(M2xM1)=det(M2)·det(M1)）。
//           编译器已证（三平台）：未跑，由收口方登记。
// 修订历史：v1.0.0 2026-11-17 首版（R24 派单 · T2-1 LGF Math 仿射变换族）
//==============================================================================

FUNCTION FC_DL_Affine2DCompose : BOOL
VAR_INPUT
    afM1 : ARRAY[0..2, 0..2] OF LREAL;      // 先施加的变换矩阵 M1 [无量纲+用户单位混合]，行主序 / First-applied transform matrix M1, row-major
    afM2 : ARRAY[0..2, 0..2] OF LREAL;      // 后施加的变换矩阵 M2 [无量纲+用户单位混合]，行主序 / Second-applied transform matrix M2, row-major
END_VAR
VAR_OUTPUT
    afMOut : ARRAY[0..2, 0..2] OF LREAL;    // 合成矩阵 MOut = M2 x M1 [无量纲+用户单位混合] / Composed matrix MOut = M2 times M1
    eErr   : UDINT;                         // 错误码，0 = 无错，码位 16#0001_0466 起信息级、16#0001_03B7 起故障级（分带见错误码表） / Error code, 0 = no error, band info/fault per the code table
    bError : BOOL;                          // 故障级标志，仅故障级错误置位 / Fault-class flag, set only on fault-level codes
    bValid : BOOL;                          // 结果可用标志 / Result usable flag
END_VAR
VAR
    afProd  : ARRAY[0..2, 0..2] OF LREAL;   // 乘积暂存阵（先算后检，检过才外泄） / Product staging array, checked before export
    nI      : INT;                          // 行循环索引 [—] / Row loop index
    nJ      : INT;                          // 列循环索引 [—] / Column loop index
    nK      : INT;                          // 求和循环索引 [—] / Summation loop index
    fAcc    : LREAL;                        // 点积累加器 [混合] / Dot-product accumulator
    fDet    : LREAL;                        // 合成矩阵线性块行列式 [无量纲] / Determinant of the composed linear block
    bNonFin : BOOL;                         // 非有限判定中间标志 / Non-finite detection intermediate flag
END_VAR
VAR CONSTANT
    DL_A2C_EPS     : LREAL := 1.0E-6;       // 行列式可逆性容差 [无量纲] / Determinant invertibility tolerance [dimensionless]
    DL_A2C_INF     : LREAL := 1.7976931348623157E308; // LREAL 幅值上限 / LREAL magnitude ceiling
    DL_A2C_ZERO    : LREAL := 0.0;          // 零值常量，避免裸字面量 [无量纲] / Zero constant, avoids a bare literal [dimensionless]
END_VAR

(*------------------------------------------------------------------------------
 * 段 1｜出口默认值：返回值与输出预置（安全侧 = 零矩阵）
 *      Exit defaults: return value and outputs preset, fail-safe zero matrix
 *-----------------------------------------------------------------------------*)
FC_DL_Affine2DCompose := FALSE;             // 返回值默认无效 / Return value preset invalid
FOR nI := 0 TO 2 DO
    FOR nJ := 0 TO 2 DO
        afMOut[nI, nJ] := DL_A2C_ZERO;      // 输出矩阵逐元素清零 / Output matrix cleared element-wise
    END_FOR
END_FOR
eErr   := 16#0000_0000;                     // 错误码先清零 / Error code cleared first
bError := FALSE;                            // 故障标志先清零 / Fault flag cleared first
bValid := FALSE;                            // 可用标志先清零 / Usable flag cleared first

(*------------------------------------------------------------------------------
 * 段 2｜输入非有限闸：两片矩阵任一元素 NaN/Inf 即拒绝（R79 双侧幅值判）
 *      Input non-finite gate over both matrices
 *-----------------------------------------------------------------------------*)
bNonFin := FALSE;                           // 非有限标志预清零 / Non-finite flag pre-cleared
FOR nI := 0 TO 2 DO
    FOR nJ := 0 TO 2 DO
        IF (afM1[nI, nJ] <> afM1[nI, nJ]) OR (ABS(afM1[nI, nJ]) > DL_A2C_INF)
           OR (afM2[nI, nJ] <> afM2[nI, nJ]) OR (ABS(afM2[nI, nJ]) > DL_A2C_INF) THEN
            bNonFin := TRUE;                // 命中非有限元素 / Non-finite element hit
        END_IF
    END_FOR
END_FOR
IF bNonFin THEN
    eErr   := 16#0001_03B7;                 // 故障级：输入矩阵元素非法 / Fault: illegal matrix element
    bError := TRUE;                         // 置故障标志（R45 配对） / Raise the fault flag
    bValid := FALSE;                        // 输出不可用 / Outputs unusable
    RETURN;                                 // 故障早退，输出保持零矩阵 / Early return, outputs stay zero
END_IF

(*------------------------------------------------------------------------------
 * 段 3｜矩阵合成：MOut = M2 x M1，完整 3x3 乘法（第三行照算不判定）
 *      Matrix composition, full 3x3 multiplication
 *-----------------------------------------------------------------------------*)
FOR nI := 0 TO 2 DO
    FOR nJ := 0 TO 2 DO
        fAcc := DL_A2C_ZERO;                // 点积累加器清零 / Accumulator cleared
        FOR nK := 0 TO 2 DO
            fAcc := fAcc + afM2[nI, nK] * afM1[nK, nJ]; // 行乘列累加 / Row-times-column accumulation
        END_FOR
        afProd[nI, nJ] := fAcc;             // 暂存乘积元素 / Stage the product element
    END_FOR
END_FOR

(*------------------------------------------------------------------------------
 * 段 4｜结果非有限复检：大坐标乘大缩放可能溢出（复用 03B7，R90）
 *      Result non-finite recheck, code reused per R90
 *-----------------------------------------------------------------------------*)
bNonFin := FALSE;                           // 非有限标志复清 / Non-finite flag re-cleared
FOR nI := 0 TO 2 DO
    FOR nJ := 0 TO 2 DO
        IF (afProd[nI, nJ] <> afProd[nI, nJ]) OR (ABS(afProd[nI, nJ]) > DL_A2C_INF) THEN
            bNonFin := TRUE;                // 命中非有限结果 / Non-finite result hit
        END_IF
    END_FOR
END_FOR
IF bNonFin THEN
    eErr   := 16#0001_03B7;                 // 故障级：结果溢出复用输入非法码（R90） / Fault: overflow, code reused per R90
    bError := TRUE;                         // 置故障标志 / Raise the fault flag
    bValid := FALSE;                        // 输出不可用 / Outputs unusable
    RETURN;                                 // 故障早退，输出保持零矩阵 / Early return, outputs stay zero
END_IF

(*------------------------------------------------------------------------------
 * 段 5｜可逆性校验：线性块行列式 |det| < 容差 → 信息级降级照常输出
 *      Invertibility check, info-level degradation with result exported
 *-----------------------------------------------------------------------------*)
fDet := afProd[0, 0] * afProd[1, 1] - afProd[0, 1] * afProd[1, 0]; // 线性块行列式 [无量纲] / Linear-block determinant
IF ABS(fDet) < DL_A2C_EPS THEN
    eErr := 16#0001_0466;                   // 信息级：合成变换不可逆（不置 bError） / Info: composed transform not invertible, no fault flag
END_IF

(*------------------------------------------------------------------------------
 * 段 6｜出口：检验通过后放行乘积阵
 *      Exit: staged product exported after checks
 *-----------------------------------------------------------------------------*)
FOR nI := 0 TO 2 DO
    FOR nJ := 0 TO 2 DO
        afMOut[nI, nJ] := afProd[nI, nJ];   // 暂存阵外泄 / Staged array exported
    END_FOR
END_FOR
bValid := TRUE;                             // 结果可用（含 0466 降级情形） / Result usable, including the degraded case
FC_DL_Affine2DCompose := TRUE;              // 返回 TRUE = 合成有效 / Return TRUE = composition valid
END_FUNCTION

(* ---- FC_DL_Affine2DInvert.st ---- *)
//==============================================================================
// 函数：FC_DL_Affine2DInvert ｜ 中文名称：二维仿射变换矩阵求逆
// 所属子库：DL_MathData ｜ 版本：v1.0.0 ｜ 兼容：CODESYS V3.5+ / TwinCAT 3 / 汇川 InoProShop
// 功能描述：3x3 仿射矩阵求逆——线性块取 2x2 伴随/行列式法，平移列按
//           t' = -A^(-1) x t 反算；点变换约定沿用本库 p' = M x p（列向量
//           右乘、行主序存储）。与 FC_DL_Affine2DCompose / FC_DL_Affine2DApply
//           构成定义-应用-逆三元闭环。与 Compose 的「不可逆降级照算」策略
//           分立：本件不可逆时输出全零矩阵，禁止半逆残阵外泄（半逆会被
//           下游点应用件当成有效映射，标定链错位难查）。库内已有
//           FC_DL_Matrix3Inverse，但其行列式含第三行，与仿射语义（第三行
//           恒为 0/0/1）不等价，按「库内委托须等价」纪律不委托、就地实现。
// 开源溯源 (Origin)：道莅 clean-room 防御性实现（仅借 LGF 分类事实/参数域/行为定义，零代码行与符号名复制）
// 单位表：矩阵线性块元素[无量纲]（旋转/缩放/剪切）/ 平移列元素[用户单位] / 行列式[无量纲]
// 错误码表：16#0001_046F 信息级（线性块奇异 |det| 小于相对判据，不可逆，
//           输出全零矩阵，不置 bError）/ 16#0001_0470 预留禁用（不得挪用）/
//           16#0001_03BD 故障级（任一输入元素非有限，或求逆结果非有限
//           溢出，置 bError，输出全零矩阵）/ 16#0001_03BE 预留禁用（不得挪用）
// 状态机：N/A——纯函数无顺序状态机，无 CASE 可写，非法状态不可能出现，以头注释说明替代 ELSE 兜底
// 边界行为：① 任一输入元素非有限（NaN 用自反判 x <> x，Inf 用幅值上限
//           兜底，R79）→ 故障 03BD、afMInv 全 0、bValid := FALSE；
//           ② |det| 小于等于 fDetEps 乘线性块最大绝对值平方（相对判据，
//           R13 Matrix3Inverse 口径）→ 信息 046F、afMInv 全 0、bValid :=
//           FALSE——不可逆禁止半逆外泄，与 Compose 降级照算策略分立；
//           ③ 第三行不参与求逆（R90 家族）：行列式与逆只按 2x2 线性块
//           加平移列计算，输出第三行按输入第三行原样回填，不做 0/0/1
//           校验（偏差提示职责归 Apply 侧，本件不重复占码位）；
//           ④ fDetEps 非正 → 回退默认 1.0E-6（容差引脚自愈，不置错）；
//           ⑤ 求逆结果非有限（大坐标乘大缩放溢出）→ 复用 03BD（R90：
//           与输入非法共用「矩阵数据不可信」语义，现有输出组合不可观测
//           出独立信息，不新占码位）、afMInv 全 0；
//           ⑥ 安全侧 = 故障与不可逆路径输出全零矩阵而非原矩阵或残阵；
//           ⑦ 失能清零不适用（纯函数无使能闸，非法输入即故障早退）。
// 修订历史：v1.0.0 2026-11-17 首版（R25 派单 · §4.1）
//==============================================================================
FUNCTION FC_DL_Affine2DInvert : BOOL
VAR_INPUT
    afM     : ARRAY[0..2, 0..2] OF LREAL;   // 待求逆仿射矩阵 M [无量纲+用户单位混合]，行主序 / Affine matrix M to invert, row-major
    fDetEps : LREAL := 1.0E-6;              // 相对奇异判据 [无量纲]，非正回退默认 / Relative singularity threshold, non-positive falls back to default
END_VAR
VAR_OUTPUT
    afMInv  : ARRAY[0..2, 0..2] OF LREAL;   // 逆矩阵 M^(-1) [无量纲+用户单位混合]，失败时全 0 / Inverse matrix, all zero on failure
    fDet    : LREAL;                        // 线性块行列式 [无量纲] / Determinant of the linear block
    eErr    : UDINT;                        // 错误码，0 = 无错，码位 16#0001_046F 起信息级、16#0001_03BD 起故障级（分带见错误码表） / Error code, 0 = no error, band info/fault per the code table
    bError  : BOOL;                         // 故障级标志，仅故障级错误置位 / Fault-class flag, set only on fault-level codes
    bValid  : BOOL;                         // 结果可用标志，不可逆与非有限路径显式 FALSE / Result usable flag, explicit FALSE on singular and non-finite paths
END_VAR
VAR
    nI      : INT;                          // 行循环索引 [—] / Row loop index
    nJ      : INT;                          // 列循环索引 [—] / Column loop index
    fMaxAbs : LREAL;                        // 线性块元素绝对值最大值 [无量纲] / Max absolute value of the linear block
    fAbsK   : LREAL;                        // 当前元素绝对值暂存 [无量纲] / Absolute value of the current element
    fEpsEff : LREAL;                        // 生效奇异判据 [无量纲] / Effective singularity threshold
    fInv00  : LREAL;                        // 逆线性块 (0,0) 元素暂存 [无量纲] / Inverse linear block element (0,0)
    fInv01  : LREAL;                        // 逆线性块 (0,1) 元素暂存 [无量纲] / Inverse linear block element (0,1)
    fInv10  : LREAL;                        // 逆线性块 (1,0) 元素暂存 [无量纲] / Inverse linear block element (1,0)
    fInv11  : LREAL;                        // 逆线性块 (1,1) 元素暂存 [无量纲] / Inverse linear block element (1,1)
    fInv02  : LREAL;                        // 逆平移列 x 分量暂存 [用户单位] / Inverse translation x component
    fInv12  : LREAL;                        // 逆平移列 y 分量暂存 [用户单位] / Inverse translation y component
    bNonFin : BOOL;                         // 非有限判定中间标志 / Non-finite detection intermediate flag
END_VAR
VAR CONSTANT
    DL_A2I_CODE_INFO_1 : UDINT := 16#0001_046F;   // 信息级槽 1（线性块奇异） / info slot 1
    DL_A2I_CODE_INFO_2 : UDINT := 16#0001_0470;   // 预留禁用（不得挪用） / reserved, do not use
    DL_A2I_CODE_FLT_1  : UDINT := 16#0001_03BD;   // 故障级槽 1（输入元素非有限） / fault slot 1
    DL_A2I_CODE_FLT_2  : UDINT := 16#0001_03BE;   // 预留禁用（不得挪用） / reserved, do not use
    DL_A2I_EPS_DEF : LREAL := 1.0E-6;               // 默认相对奇异判据 [无量纲] / Default relative singularity threshold [dimensionless]
    DL_A2I_INF     : LREAL := 1.7976931348623157E308; // LREAL 幅值上限，Inf 判据 / LREAL magnitude ceiling, Inf criterion
    DL_A2I_ZERO    : LREAL := 0.0;                  // 零值常量，避免裸字面量 [无量纲] / Zero constant, avoids a bare literal [dimensionless]
END_VAR

(*------------------------------------------------------------------------------
 * 段 1｜出口默认值先行：全零矩阵 + 无错 + 不可用（先写后算，任何早退路径出口确定）
 *----------------------------------------------------------------------------*)
FOR nI := 0 TO 2 DO
    FOR nJ := 0 TO 2 DO
        afMInv[nI, nJ] := DL_A2I_ZERO;         // 逆矩阵默认全零 / default all-zero inverse
    END_FOR
END_FOR
fDet   := DL_A2I_ZERO;                         // 行列式默认零 / determinant defaults to zero
eErr   := 16#0000_0000;                        // 错误码默认无错 / error code defaults to none
bError := FALSE;                               // 故障标志默认清除 / fault flag cleared
bValid := FALSE;                               // 可用标志默认不可用，算完并检过才置位 / usable flag FALSE until computed and checked

(*------------------------------------------------------------------------------
 * 段 2｜输入非有限全阵扫描（9 元素逐个：NaN 自反判 + Inf 幅值上限判，R79）
 *----------------------------------------------------------------------------*)
bNonFin := FALSE;                              // 非有限标志复位 / reset non-finite flag
FOR nI := 0 TO 2 DO
    FOR nJ := 0 TO 2 DO
        IF (afM[nI, nJ] <> afM[nI, nJ]) OR (ABS(afM[nI, nJ]) >= DL_A2I_INF) THEN
            bNonFin := TRUE;                   // 发现非有限元素 / non-finite element found
        END_IF
    END_FOR
END_FOR
IF bNonFin THEN
    eErr   := DL_A2I_CODE_FLT_1;               // 故障级：任一输入元素非有限 / fault: non-finite input element
    bError := TRUE;                            // 故障级必置 bError（R45 配对）/ fault-class pairs with bError
    bValid := FALSE;                           // 输出不可用 / outputs unusable
    FC_DL_Affine2DInvert := FALSE;             // 返回值 = 可用标志同口径 / return mirrors bValid
    RETURN;
END_IF

(*------------------------------------------------------------------------------
 * 段 3｜线性块行列式与相对奇异判据（第三行不参与，R90 家族）
 *----------------------------------------------------------------------------*)
fDet := afM[0, 0] * afM[1, 1] - afM[0, 1] * afM[1, 0];  // 2x2 线性块行列式 / 2x2 linear block determinant
fMaxAbs := ABS(afM[0, 0]);                     // 最大绝对值种子：m00 / seed max with m00
fAbsK := ABS(afM[0, 1]);                       // m01 绝对值 / absolute of m01
IF fAbsK > fMaxAbs THEN fMaxAbs := fAbsK; END_IF
fAbsK := ABS(afM[1, 0]);                       // m10 绝对值 / absolute of m10
IF fAbsK > fMaxAbs THEN fMaxAbs := fAbsK; END_IF
fAbsK := ABS(afM[1, 1]);                       // m11 绝对值 / absolute of m11
IF fAbsK > fMaxAbs THEN fMaxAbs := fAbsK; END_IF
fEpsEff := fDetEps;                            // 生效判据先取引脚 / effective threshold from pin
IF fEpsEff <= DL_A2I_ZERO THEN
    fEpsEff := DL_A2I_EPS_DEF;                 // 非正回退默认判据 / non-positive falls back to default
END_IF
IF ABS(fDet) <= fEpsEff * fMaxAbs * fMaxAbs THEN
    eErr   := DL_A2I_CODE_INFO_1;              // 信息级：线性块奇异，不可逆 / info: singular linear block, not invertible
    bError := FALSE;                           // 信息级不置 bError（R45/R101）/ info never raises bError
    bValid := FALSE;                           // 逆矩阵不可用，禁止半逆外泄 / inverse unusable, no half-inverse leak
    FC_DL_Affine2DInvert := FALSE;             // 返回值同口径 / return mirrors bValid
    RETURN;
END_IF

(*------------------------------------------------------------------------------
 * 段 4｜2x2 伴随求逆 + 平移列反算 t' = -A^(-1) x t（除子 fDet 已由段 3 保证非零）
 *----------------------------------------------------------------------------*)
fInv00 :=  afM[1, 1] / fDet;                   // A^(-1)(0,0) = m11/det / inverse element
fInv01 := -afM[0, 1] / fDet;                   // A^(-1)(0,1) = -m01/det / inverse element
fInv10 := -afM[1, 0] / fDet;                   // A^(-1)(1,0) = -m10/det / inverse element
fInv11 :=  afM[0, 0] / fDet;                   // A^(-1)(1,1) = m00/det / inverse element
fInv02 := -(fInv00 * afM[0, 2] + fInv01 * afM[1, 2]);  // 逆平移列 x = -(A^(-1) x t)_x / inverse translation x
fInv12 := -(fInv10 * afM[0, 2] + fInv11 * afM[1, 2]);  // 逆平移列 y = -(A^(-1) x t)_y / inverse translation y

(*------------------------------------------------------------------------------
 * 段 5｜结果非有限复检（溢出复用 03BD，见边界行为⑤）后装配输出
 *----------------------------------------------------------------------------*)
IF (fInv00 <> fInv00) OR (fInv01 <> fInv01) OR (fInv10 <> fInv10) OR (fInv11 <> fInv11)
   OR (fInv02 <> fInv02) OR (fInv12 <> fInv12)
   OR (ABS(fInv00) >= DL_A2I_INF) OR (ABS(fInv01) >= DL_A2I_INF)
   OR (ABS(fInv10) >= DL_A2I_INF) OR (ABS(fInv11) >= DL_A2I_INF)
   OR (ABS(fInv02) >= DL_A2I_INF) OR (ABS(fInv12) >= DL_A2I_INF) THEN
    FOR nI := 0 TO 2 DO
        FOR nJ := 0 TO 2 DO
            afMInv[nI, nJ] := DL_A2I_ZERO;     // 溢出路径安全侧：全零矩阵 / overflow path safe side: all-zero
        END_FOR
    END_FOR
    eErr   := DL_A2I_CODE_FLT_1;               // 故障级：求逆结果非有限溢出 / fault: non-finite inverse result
    bError := TRUE;                            // 故障级必置 bError（R45 配对）/ fault-class pairs with bError
    bValid := FALSE;                           // 输出不可用 / outputs unusable
    FC_DL_Affine2DInvert := FALSE;             // 返回值同口径 / return mirrors bValid
    RETURN;
END_IF

(*------------------------------------------------------------------------------
 * 段 6｜装配输出：线性块 + 平移列 + 第三行原样回填（边界行为③）
 *----------------------------------------------------------------------------*)
afMInv[0, 0] := fInv00;                        // 逆线性块 (0,0) / inverse element
afMInv[0, 1] := fInv01;                        // 逆线性块 (0,1) / inverse element
afMInv[0, 2] := fInv02;                        // 逆平移列 x / inverse translation x
afMInv[1, 0] := fInv10;                        // 逆线性块 (1,0) / inverse element
afMInv[1, 1] := fInv11;                        // 逆线性块 (1,1) / inverse element
afMInv[1, 2] := fInv12;                        // 逆平移列 y / inverse translation y
afMInv[2, 0] := afM[2, 0];                     // 第三行原样回填，不校验 / third row copied verbatim, unchecked
afMInv[2, 1] := afM[2, 1];                     // 第三行原样回填，不校验 / third row copied verbatim, unchecked
afMInv[2, 2] := afM[2, 2];                     // 第三行原样回填，不校验 / third row copied verbatim, unchecked
eErr   := 16#0000_0000;                        // 无错出口 / no-error exit
bError := FALSE;                               // 无故障 / no fault
bValid := TRUE;                                // 逆矩阵可用 / inverse usable
FC_DL_Affine2DInvert := TRUE;                  // 返回值 = 可用标志 / return mirrors bValid
END_FUNCTION

(* ---- FC_DL_AffineTransformPoint.st ---- *)
(*
    FC_DL_AffineTransformPoint —— 2D 仿射点变换
    ------------------------------------------------------------------
    分类      : DL_MathData / Transform
    前缀      : FC_DL_
    版本      : 1.0.0
    溯源      : T2-1 LGF · Math（源矩阵明列「仿射变换组合族待挖」；只借该族归属
                Math 的分类事实）；旋转 / 缩放 / 平移的合成顺序为本库自有规格，
                角度归一式的工程写法、码位与错误分级 100% 自有；
                clean-room 重写，未复制任何闭源厂商源码，参考实现仅限 MIT/Apache 许可
    平台      : 纯 IEC 61131-3，CODESYS V3.5+ / TwinCAT 3 / InoProShop 通用
    作者      : 道莅代码库 · PLC编程专家（R18）
    ------------------------------------------------------------------
    功能说明  : 单次完成「绕原点旋转 → 各轴缩放 → 平移」的合成，输出变换后坐标。
                现场语义：视觉像素坐标到机械 mm 坐标（含相机安装角偏差）、纠偏平台
                坐标映射、印刷套准偏移换算；
                角度归一用「减 360 乘整数商」单算式路径，不用循环也不用取余
                （浮点取余在三平台行为不一致）；三角函数直接调用内建 SIN / COS，
                绝不重实现（T0 判据 2）；
                缩放为 0 使变换不可逆，按故障拒绝并原值回送，绝不返回被压平的点；
                输入与中间结果双向非有限复检，1e38 量级缩放乘大坐标的溢出能被抓住。
    错误码    : 16#0001_0241 旋转角超正负 360 度已归一——信息级，正常防御
                16#0001_0242 预留禁用（信息级，不得挪用）
                16#0001_0318 缩放因子为 0（变换不可逆）——故障级，返回原点值
                16#0001_0319 输入或中间结果非有限（NaN / 正负 INF / 溢出）——故障级，输出 0
                16#0001_031A 预留禁用（故障级，不得挪用）
    码位总账  : 16#0001_0241 用 / 16#0001_0242 预留 ｜ 16#0001_0318 用 / 16#0001_0319 用 / 16#0001_031A 预留
    状态机    : N/A —— 纯函数无顺序状态机，无 CASE 可写，非法状态不可能出现
    采样约定  : 纯组合函数，无定时器、无内部驻留状态；变换参数由调用方保证在同一
                标定批次内恒定（本库统一约定：标定参数只在停机态下发）。
    修订记录  : 2026-11-16 v1.0.0 首次入库（R18）
*)
FUNCTION FC_DL_AffineTransformPoint : BOOL
VAR_INPUT
    fX       : REAL := 0.0;                    // 源点 X [用户单位] / source point X [user unit]
    fY       : REAL := 0.0;                    // 源点 Y [用户单位] / source point Y [user unit]
    fRotDeg  : REAL := 0.0;                    // 旋转角，正为逆时针 [度]，范围 -720.0~720.0 / rotation angle, positive counter clockwise [deg], range -720.0~720.0
    fScaleX  : REAL := 1.0;                    // X 缩放比 [比值]，范围 0.001~1000.0，禁 0 / X scale ratio [ratio], range 0.001~1000.0, zero forbidden
    fScaleY  : REAL := 1.0;                    // Y 缩放比 [比值]，范围 0.001~1000.0，禁 0 / Y scale ratio [ratio], range 0.001~1000.0, zero forbidden
    fTx      : REAL := 0.0;                    // X 平移量 [用户单位] / X translation [user unit]
    fTy      : REAL := 0.0;                    // Y 平移量 [用户单位] / Y translation [user unit]
END_VAR
VAR_OUTPUT
    fOutX  : REAL;                             // 变换后 X [用户单位] / transformed X [user unit]
    fOutY  : REAL;                             // 变换后 Y [用户单位] / transformed Y [user unit]
    eErr   : UDINT;                            // 错误码，0=正常 / error id, 0=ok
    bError : BOOL;                             // 故障标志，eErr 为故障级时 TRUE / error flag, TRUE on fault-level eErr
    bValid : BOOL;                             // 结果是否可用 / result usable flag
END_VAR
VAR
    fAngNorm : REAL;                           // 归一后角度 [度]，范围 0~360 / normalised angle [deg], range 0~360
    fRad     : REAL;                           // 归一后角度换算的弧度 [弧度] / normalised angle in radians [rad]
    fCos     : REAL;                           // 余弦值，范围 -1.0~1.0 [无量纲] / cosine value, range -1.0~1.0 [dimensionless]
    fSin     : REAL;                           // 正弦值，范围 -1.0~1.0 [无量纲] / sine value, range -1.0~1.0 [dimensionless]
    fXRot    : REAL;                           // 旋转后 X [用户单位] / X after rotation [user unit]
    fYRot    : REAL;                           // 旋转后 Y [用户单位] / Y after rotation [user unit]
    fXScaled : REAL;                           // 缩放后 X [用户单位] / X after scaling [user unit]
    fYScaled : REAL;                           // 缩放后 Y [用户单位] / Y after scaling [user unit]
    fQuot    : REAL;                           // 角度除以 360 的整数商中间量 [无量纲] / integer quotient of the angle divided by 360 [dimensionless]
    bNonFin  : BOOL;                           // 非有限判定中间标志 / non-finite detection intermediate flag
END_VAR
VAR CONSTANT
    DL_AFF_EPS        : REAL := 1.0E-6;        // 浮点判等容差 [无量纲] / float equality tolerance [dimensionless]
    DL_AFF_INF_GUARD  : REAL := 4.0E38;        // 非有限幅值判定阈值，高于 REAL 最大有限值 [用户单位] / non-finite magnitude guard above the largest finite REAL [user unit]
    DL_AFF_FULL_DEG   : REAL := 360.0;         // 一整圈角度 [度] / one full turn [deg]
    DL_AFF_DEG2RAD    : REAL := 0.017453292519943295; // 度转弧度系数 [弧度每度] / degree to radian factor [rad per deg]
    DL_AFF_ZERO       : REAL := 0.0;           // 零值常量，避免裸字面量 [无量纲] / zero constant, avoids a bare literal [dimensionless]
    DL_AFF_TWO        : REAL := 2.0;           // 除数二，用于半圆判定 [无量纲] / divisor two, used by the half turn check [dimensionless]
END_VAR

// 段 1｜返回值与输出预置 / segment 1, preset return value and outputs
FC_DL_AffineTransformPoint := FALSE;           // 故障缺省返回 FALSE / fault default returns FALSE
fOutX := DL_AFF_ZERO;                          // 输出 X 预置 0 / preset X to zero
fOutY := DL_AFF_ZERO;                          // 输出 Y 预置 0 / preset Y to zero
eErr := 0;                                     // 预置无错误 / preset no error
bError := FALSE;                               // 预置无故障 / preset no fault
bValid := FALSE;                               // 预置结果不可用 / preset unusable

// 段 2｜输入非有限闸：任一输入 NaN 或正负 INF 即拒绝 / segment 2, input non-finite gate
bNonFin := (fX <> fX) OR (fX > DL_AFF_INF_GUARD) OR (fX < -DL_AFF_INF_GUARD)
        OR (fY <> fY) OR (fY > DL_AFF_INF_GUARD) OR (fY < -DL_AFF_INF_GUARD)
        OR (fRotDeg <> fRotDeg) OR (fRotDeg > DL_AFF_INF_GUARD) OR (fRotDeg < -DL_AFF_INF_GUARD)
        OR (fTx <> fTx) OR (fTx > DL_AFF_INF_GUARD) OR (fTx < -DL_AFF_INF_GUARD)
        OR (fTy <> fTy) OR (fTy > DL_AFF_INF_GUARD) OR (fTy < -DL_AFF_INF_GUARD); // 平移与角度同样检查 / translation and angle are checked the same way
IF bNonFin THEN
    eErr := 16#0001_0319;                      // 输入非有限故障码 / non-finite input fault id
    bError := TRUE;                            // 置故障标志 / raise the error flag
    RETURN;                                    // 故障级提前返回，输出保持 0 / early return on fault, outputs stay zero
END_IF

// 段 3｜缩放闸：缩放为 0 使变换不可逆，原值回送并拒绝 / segment 3, zero scale gate
IF (ABS(fScaleX) < DL_AFF_EPS) OR (ABS(fScaleY) < DL_AFF_EPS) THEN
    eErr := 16#0001_0318;                      // 缩放为零故障码 / zero scale fault id
    bError := TRUE;                            // 置故障标志 / raise the error flag
    fOutX := fX;                               // 原值回送 X，便于上层诊断 / return the original X so the caller can diagnose
    fOutY := fY;                               // 原值回送 Y / return the original Y
    RETURN;                                    // 故障级提前返回 / early return on fault
END_IF

// 段 4｜角度归一：减 360 乘以整数商，单算式路径，不用循环也不用取余 / segment 4, angle normalisation
fAngNorm := fRotDeg;                           // 默认沿用输入角 / default to the input angle
IF ABS(fRotDeg) > DL_AFF_FULL_DEG THEN
    fQuot := TRUNC(fRotDeg / DL_AFF_FULL_DEG); // 整数商（向零截断，除数为常量 360 恒非零）/ integer quotient, truncated toward zero, the divisor is the constant 360
    fAngNorm := fRotDeg - DL_AFF_FULL_DEG * fQuot; // 单算式归一，残差落在正负 360 内 / single expression normalisation, the residual stays within plus or minus 360
    eErr := 16#0001_0241;                      // 归一提示（信息级不置故障）/ normalisation hint, info level never raises a fault
END_IF

// 段 5｜三角函数：直接调内建，绝不重实现 / segment 5, trigonometric functions are built-in calls only
fRad := fAngNorm * DL_AFF_DEG2RAD;             // 度转弧度 / degrees to radians
fCos := COS(fRad);                             // 余弦 [无量纲] / cosine [dimensionless]
fSin := SIN(fRad);                             // 正弦 [无量纲] / sine [dimensionless]

// 段 6｜旋转 → 缩放 → 平移 合成 / segment 6, rotation then scaling then translation
fXRot := fX * fCos - fY * fSin;                // 旋转后 X / X after rotation
fYRot := fX * fSin + fY * fCos;                // 旋转后 Y / Y after rotation
fXScaled := fXRot * fScaleX;                   // 各轴缩放 X / per axis scaling on X
fYScaled := fYRot * fScaleY;                   // 各轴缩放 Y / per axis scaling on Y
fOutX := fXScaled + fTx;                       // 叠加 X 平移 / add the X translation
fOutY := fYScaled + fTy;                       // 叠加 Y 平移 / add the Y translation

// 段 7｜结果非有限复检：大缩放乘大坐标可能溢出 / segment 7, result non-finite recheck
bNonFin := (fOutX <> fOutX) OR (fOutX > DL_AFF_INF_GUARD) OR (fOutX < -DL_AFF_INF_GUARD)
        OR (fOutY <> fOutY) OR (fOutY > DL_AFF_INF_GUARD) OR (fOutY < -DL_AFF_INF_GUARD); // 结果溢出判定 / result overflow check
IF bNonFin THEN
    fOutX := DL_AFF_ZERO;                      // 溢出即输出 0 / overflow yields zero
    fOutY := DL_AFF_ZERO;                      // 溢出即输出 0 / overflow yields zero
    eErr := 16#0001_0319;                      // 结果非有限故障码 / non-finite result fault id
    bError := TRUE;                            // 置故障标志 / raise the error flag
    RETURN;                                    // 故障级提前返回 / early return on fault
END_IF

// 段 8｜出口 / segment 8, exit
bValid := TRUE;                                // 结果可用 / the result is usable
FC_DL_AffineTransformPoint := TRUE;            // 变换成功 / the transform succeeded
END_FUNCTION

(* ---- FC_DL_AkimaInterp1D.st ---- *)
(*
  道莅工业代码库 | DL_MathData | FC_DL_AkimaInterp1D
  版本: 1.0.0 | 日期: 2026-11-23 | 轮次: R75
  开源溯源: self-cleanroom（无外部来源；Akima 1970 抗振荡插值为公开算法，
            本件独立实现，零代码行复制）
  功能: Akima 一维插值（显式点数入参防 VLA）——5 点及以上走完整 Akima
        切线加权（端部斜率外推两支），2~4 点回落线性插值；查询点越界钳端点。
  兼容性: CODESYS 3.5 / TwinCAT 3 / 汇川 InoProShop；仅依赖标准 ABS/SQRT，零厂商私有库
  接口: 输入查询点 fX、节点表 aX/aY（固定上界 ARRAY[1..100] OF REAL）、
        uPointCnt（1..200，内部钳位 [2,100]）；返回值 TRUE=已执行；
        输出 fY（越界钳端点值）、bValid、eErr。纯函数：无内部状态。
  码表: 16#0001_0500 故障级：节点表非法（含非有限值或未严格升序，或查询点 NaN）
        码段说明：0001 段 03xx 故障子带已满（03FF 已占用），启用 05xx 扩展域闸子带，
        0500 槽经全库实扫空闲。
  边界: ① uPointCnt 先钳位 [2,100]（R75 显式点数字段口径），钳位后 < 2 不可能，
        表非法仅由升序破坏/非有限/查询 NaN 触发；
        ② 段斜率除法分母由升序闸（节点差 > EPS）证明 > 0；
        ③ Akima 切线权重分母 (w1+w2) = 0 时回落两邻段斜率均值（算法标准防除零）；
        ④ 端部外推斜率 m0/m-1/mn/mn+1 需 n >= 4，本件以 n >= 5 进 Akima 路径闸住；
        ⑤ 全部输出在所有路径（含提前返回）赋值；⑥ 零全局耦合。
  邻件比对: Lagrange/Hermite/CubicSpline（多项式样条族 vs 本件 Akima 抗振荡切线族）。
  修订历史: 2026-11-23 v1.0.0 R75 首版（复杂件批 B2 · C09）
*)

FUNCTION FC_DL_AkimaInterp1D : BOOL
VAR_INPUT
    fX        : REAL;                     // 查询点横坐标 [x 单位] | Query abscissa
    aX        : ARRAY[1..100] OF REAL;    // 节点横坐标表（严格升序）[x 单位] | Node abscissae, strictly ascending
    aY        : ARRAY[1..100] OF REAL;    // 节点纵坐标表 [y 单位] | Node ordinates
    uPointCnt : UINT := 5;                // 有效点数，内部钳位 [2,100] [点] | Valid point count, clamped internally
END_VAR
VAR_OUTPUT
    fY     : REAL;                        // 插值结果（越界钳端点值）[y 单位] | Interpolated result, clamped at bounds
    bValid : BOOL;                        // 本次计算有效 [-] | Computation valid
    eErr   : UDINT;                       // 错误码，0 = 无错 | Error code, 0 = none
END_VAR
VAR
    nI      : INT;                        // 钳位后点数 [点] | Clamped point count
    i       : INT;                        // 循环游标 | Loop cursor
    iSeg    : INT;                        // 所在段左节点序号 | Segment left knot index
    bTabOk  : BOOL;                       // 表合法当拍量 [-] | Table legality this call
    bAkima  : BOOL;                       // Akima 路径标志（n >= 5）[-] | Akima path flag
    fQ      : REAL;                       // 钳界后查询点 [x 单位] | Clamped query point
    fDx     : REAL;                       // 段宽 [x 单位] | Segment width
    fTParam : REAL;                       // 段内归一化参数 t ∈ [0, 1] [-] | Normalized parameter in segment
    fT2     : REAL;                       // t 的平方 [-] | t squared
    fT3     : REAL;                       // t 的立方 [-] | t cubed
    w1      : REAL;                       // Akima 权重 |m_{i+1}-m_i| [-] | Akima weight upper
    w2      : REAL;                       // Akima 权重 |m_{i-1}-m_{i-2}| [-] | Akima weight lower
    aM      : ARRAY[1..103] OF REAL;      // 段斜率数组（含端部外拓 m_-1..m_n+1，下标偏移 +2）[y/x] | Segment slopes with two-sided extension, index offset +2
    aTang      : ARRAY[1..100] OF REAL;      // 节点切线数组 [y/x] | Knot tangents
END_VAR
VAR CONSTANT
    DL_AKI_EPS : REAL := 1.0E-6;          // 升序判据容差（节点最小间距）[x 单位] | Ascending tolerance
    DL_AKI_ERR : UDINT := 16#0001_0500;   // 节点表非法码 | Illegal table code
END_VAR

(* —— 段 0：输出缺省全赋值（全路径覆盖） —— *)
fY := 0.0;                                // 结果预置零 / Result preset zero
bValid := FALSE;                          // 有效标志预置 / Valid preset FALSE
eErr := 0;                                // 错误码缺省 / Error default
FC_DL_AkimaInterp1D := TRUE;              // 返回值：TRUE = 已执行 / Result: TRUE = executed

(* —— 段 1：点数钳位与表合法性闸（R75 显式点数字段口径） —— *)
nI := UINT_TO_INT(uPointCnt);             // 点数转整型 / Point count to INT
IF nI < 2 THEN
    nI := 2;                              // 下限钳 2（至少两点） / Clamp lower to 2
END_IF
IF nI > 100 THEN
    nI := 100;                            // 上限钳 100（数组容量） / Clamp upper to 100
END_IF
bTabOk := (fX = fX);                      // 查询点 NaN 自反判 / Query NaN self-reflex check
IF bTabOk THEN
    FOR i := 1 TO nI DO
        IF (aX[i] <> aX[i]) OR (aY[i] <> aY[i]) THEN
            bTabOk := FALSE;              // 节点值非有限 / Node value non-finite
        END_IF
    END_FOR
END_IF
IF bTabOk THEN
    FOR i := 1 TO (nI - 1) DO
        IF (aX[i + 1] - aX[i]) <= DL_AKI_EPS THEN
            bTabOk := FALSE;              // 严格升序被破坏（含重合节点） / Strict ascending violated
        END_IF
    END_FOR
END_IF
IF NOT bTabOk THEN
    eErr := DL_AKI_ERR;                   // 表非法码 / Illegal table code
    RETURN;                               // 提前返回：输出已全赋值 / Early return, outputs assigned
END_IF

(* —— 段 2：查询点钳界 —— *)
fQ := fX;                                 // 查询点暂存 / Query staging
IF fQ < aX[1] THEN
    fQ := aX[1];                          // 下界钳首节点 / Clamp to first knot
END_IF
IF fQ > aX[nI] THEN
    fQ := aX[nI];                         // 上界钳末节点 / Clamp to last knot
END_IF
bAkima := nI >= 5;                        // 5 点及以上走 Akima（端部外拓需 n >= 4） / Akima path for n >= 5

(* —— 段 3：Akima 段斜率与端部外拓 —— *)
IF bAkima THEN
    FOR i := 1 TO (nI - 1) DO
        fDx := aX[i + 1] - aX[i];         // 段宽（升序闸保证 > EPS） / Segment width, proven positive
        aM[i + 2] := (aY[i + 1] - aY[i]) / fDx;   // 段斜率 m_i 存 aM[i+2] / Segment slope, offset +2
    END_FOR
    aM[2] := 2.0 * aM[3] - aM[4];         // 端部外拓 m_0 = 2m_1 - m_2 / Extended slope m0
    aM[1] := 2.0 * aM[2] - aM[3];         // 端部外拓 m_-1 = 2m_0 - m_1 / Extended slope m-1
    aM[nI + 2] := 2.0 * aM[nI + 1] - aM[nI];       // 端部外拓 m_n = 2m_n-1 - m_n-2 / Extended slope mn
    aM[nI + 3] := 2.0 * aM[nI + 2] - aM[nI + 1];   // 端部外拓 m_n+1 = 2m_n - m_n-1 / Extended slope mn+1

    (* —— 段 4：节点切线（Akima 加权；权重和零回落均值防除零） —— *)
    FOR i := 1 TO nI DO
        w1 := ABS(aM[i + 3] - aM[i + 2]); // 权重 w1 = |m_{i+1} - m_i| / Weight from adjacent slope gap
        w2 := ABS(aM[i + 1] - aM[i]);     // 权重 w2 = |m_{i-1} - m_{i-2}| / Weight from second-adjacent gap
        IF (w1 + w2) > DL_AKI_EPS THEN
            aTang[i] := (w1 * aM[i + 1] + w2 * aM[i + 2]) / (w1 + w2);   // 加权切线（分母已闸）/ Weighted tangent, denominator gated
        ELSE
            aTang[i] := 0.5 * (aM[i + 1] + aM[i + 2]);   // 权重和零回落两邻段均值 / Fallback to mean of adjacent slopes
        END_IF
    END_FOR
END_IF

(* —— 段 5：段定位（fQ 已钳在 [aX[1], aX[nI]]，循环有界） —— *)
iSeg := 1;                                // 段定位从首段起 / Segment search from first
WHILE (iSeg < (nI - 1)) AND (fQ > aX[iSeg + 1]) DO
    iSeg := iSeg + 1;                     // 右移至目标段 / Advance to target segment
END_WHILE

(* —— 段 6：段内插值（Akima 三次 Hermite / 回落线性） —— *)
fDx := aX[iSeg + 1] - aX[iSeg];           // 段宽（升序闸保证 > EPS） / Segment width, proven positive
fTParam := (fQ - aX[iSeg]) / fDx;         // 归一化参数，分母已闸 / Normalized parameter, denominator gated
IF bAkima THEN
    fT2 := fTParam * fTParam;             // t² / t squared
    fT3 := fT2 * fTParam;                 // t³ / t cubed
    fY := aY[iSeg] * (2.0 * fT3 - 3.0 * fT2 + 1.0)
       + aY[iSeg + 1] * (3.0 * fT2 - 2.0 * fT3)
       + fDx * aTang[iSeg] * (fT3 - 2.0 * fT2 + fTParam)
       + fDx * aTang[iSeg + 1] * (fT3 - fT2);            // 三次 Hermite 基函数合成 / Cubic Hermite basis synthesis
ELSE
    fY := aY[iSeg] + fTParam * (aY[iSeg + 1] - aY[iSeg]);  // 线性回落（n < 5）/ Linear fallback
END_IF
bValid := TRUE;                           // 计算有效 / Valid

END_FUNCTION

(* ---- FC_DL_AmpDbToRatio.st ---- *)
(*
    FC_DL_AmpDbToRatio —— 幅值型分贝到线性幅值比换算
    ------------------------------------------------------------------
    分类      : DL_MathData / Log
    前缀      : FC_DL_
    版本      : 1.0.0
    溯源      : IEC 61131-3 标准语义的道莅防御性实现
                （接口语义由 IEC 61131-3 定义，内部委托平台内建 EXPT，
                  外围统一错误码 / 钳位 / 双语文档；clean-room 重写，
                  未复制任何闭源厂商源码，参考实现仅限 MIT/Apache 许可）
    平台      : 纯 IEC 61131-3，CODESYS / TwinCAT / InoProShop 通用
    作者      : 道莅代码库 · PLC编程专家（R17）
    ------------------------------------------------------------------
    功能说明  : 幅值型分贝转过线性幅值比，按 A = 10^(dB/20) 实现，指数运算委托平台内建 EXPT，
                20 为幅值型换算因子（与功率型 10 严格区分，禁混用），不重实现指数内核；
                非有限输入判为故障级 16#0001_02D0，返回 1.0（比值中性值，避免下游乘零灭信号）；
                |dB| 超 400.0 dB 硬限时按方向饱和至 1.0E20 / 1.0E-20，置信息级 16#0001_01EC；
                EXPT 结果复检非有限（部分平台溢出行为不一致）同样按方向饱和并复用 01EC；
                钳位方向：双侧饱和（dB 域 ±400.0 dB，比值域 1.0E-20 ~ 1.0E20）。
    错误码    : 16#0001_01EC dB 值超 ±400.0 dB 硬限，已按方向饱和——信息级，正常防御
                16#0001_01ED 预留禁用（信息级，不得挪用）
                16#0001_02D0 非有限输入（NaN 或 ±INF）——故障级，返回 1.0
                16#0001_02D1 预留禁用（故障级，不得挪用）
                16#0001_02D2 预留禁用（故障级，不得挪用）
    状态机    : R6 标注 N/A —— 本组件为纯函数无顺序状态机，无 CASE 可写，非法状态不可能出现，故以本节说明替代 ELSE 兜底
    修订记录  : 2026-11-16 v1.0.0 首次入库（R17）
*)
FUNCTION FC_DL_AmpDbToRatio : REAL
VAR_INPUT
    fDb : REAL; // 幅值型分贝值，建议域 −400.0~+400.0 [dB] / amplitude decibel value, suggested domain -400.0..+400.0 [dB]
END_VAR
VAR_OUTPUT
    eErr   : UDINT; // 错误码，0=正常 / error id, 0=ok
    bError : BOOL;  // 是否出错，eErr 非 0 时为 TRUE / error flag, TRUE when eErr is nonzero
    bValid : BOOL;  // 输出是否有效可用 / output valid flag
END_VAR
VAR CONSTANT
    DL_DB_AMP_DIV     : REAL := 20.0;      // 幅值型 dB 换算除子（20·log10 的逆向） [dB] / amplitude dB divisor, inverse of 20*log10 [dB]
    DL_DB_TEN         : REAL := 10.0;      // 幂运算底数 10 [无量纲] / power base 10 [dimensionless]
    DL_DB_LIMIT       : REAL := 400.0;     // dB 域双侧硬限，对应比值 10^±20 [dB] / two-sided dB hard limit, ratio 10^+/-20 [dB]
    DL_RATIO_NEUTRAL  : REAL := 1.0;       // 比值中性值（0 dB 对应值，故障缺省返回） [比] / neutral ratio (0 dB), fault default [ratio]
    DL_RATIO_MAX      : REAL := 1.0E20;    // 幅值比上限 10^20，REAL 域可表 [比] / amplitude ratio upper bound 10^20 [ratio]
    DL_RATIO_MIN      : REAL := 1.0E-20;   // 幅值比下限 10^-20，REAL 域可表 [比] / amplitude ratio lower bound 10^-20 [ratio]
    DL_REAL_INF_GUARD : LREAL := 4.0E38;   // REAL 域 ±INF 判定阈值，高于 REAL 最大有限值 3.402823E38 [无量纲] / REAL +/-INF guard above max finite REAL
END_VAR
VAR
    bNonFinite : BOOL; // 非有限（NaN 或 ±INF）判定结果 / non-finite (NaN or +/-INF) detection result
END_VAR

// 段 1｜返回值与错误状态预置 / segment 1, preset return value and error status
FC_DL_AmpDbToRatio := DL_RATIO_NEUTRAL; // 故障缺省返回 1.0 中性比值，避免下游乘零灭信号 [比] / fault default 1.0 neutral ratio, avoids killing the signal downstream [ratio]
eErr   := 0;     // 预置无错误 / preset no error
bError := FALSE; // 预置无故障 / preset no fault
bValid := FALSE; // 预置输出无效，通过非有限闸后置位 / preset invalid, set TRUE after the non-finite gate

// 段 2｜非有限防御闸 / segment 2, non-finite guard
bNonFinite := (fDb <> fDb) OR (fDb > DL_REAL_INF_GUARD) OR (fDb < -DL_REAL_INF_GUARD); // 非有限判定（NaN 自不等 + 安全幅值判 ±INF） [dB] / non-finite check (NaN by self-inequality, +/-INF by safe magnitude) [dB]
IF bNonFinite THEN
    eErr := 16#0001_02D0; // 非有限输入故障码 / non-finite input fault id
    bError := TRUE;       // 置故障标志 / raise error flag
    bValid := FALSE;      // 输出不可用 / output not usable
    RETURN;               // 故障级提前返回，保持缺省 1.0 / early return on fault, keep default 1.0
END_IF

// 段 3｜dB 域硬限双侧饱和 / segment 3, two-sided dB domain saturation
IF fDb > DL_DB_LIMIT THEN
    FC_DL_AmpDbToRatio := DL_RATIO_MAX; // 正超饱和至幅值比上限 1.0E20 [比] / positive overflow saturates to ratio upper bound 1.0E20 [ratio]
    eErr := 16#0001_01EC;               // 信息级：dB 超限已饱和，正常防御 / info level: dB exceeded the limit and saturated, normal defence
    bError := FALSE;                    // 信息级不置故障 / info level never raises fault
    bValid := TRUE;                     // 饱和值本身有效可用 / the saturated value itself is valid
    RETURN;                             // 饱和即出口，不进入幂运算 / saturation is the exit, no power computation
END_IF
IF fDb < -DL_DB_LIMIT THEN
    FC_DL_AmpDbToRatio := DL_RATIO_MIN; // 负超饱和至幅值比下限 1.0E-20 [比] / negative overflow saturates to ratio lower bound 1.0E-20 [ratio]
    eErr := 16#0001_01EC;               // 同一业务语义复用同一信息码 / same business semantics reuses the same info id
    bError := FALSE;                    // 信息级不置故障 / info level never raises fault
    bValid := TRUE;                     // 饱和值本身有效可用 / the saturated value itself is valid
    RETURN;                             // 饱和即出口，不进入幂运算 / saturation is the exit, no power computation
END_IF

// 段 4｜主体幂运算与结果复检（末段） / segment 4, main power computation and result re-check (final)
FC_DL_AmpDbToRatio := EXPT(DL_DB_TEN, fDb / DL_DB_AMP_DIV); // 域内委托内建 EXPT 计算 10^(dB/20) [比] / in-domain delegate to built-in EXPT for 10^(dB/20) [ratio]
IF (FC_DL_AmpDbToRatio <> FC_DL_AmpDbToRatio) OR (FC_DL_AmpDbToRatio > DL_RATIO_MAX) OR (FC_DL_AmpDbToRatio < DL_RATIO_MIN) THEN // 结果复检：NaN 自不等 + 双侧越界（±INF 亦被幅值界捕获） [比] / result re-check: NaN by self-inequality plus two-sided overflow, +/-INF also caught by the magnitude bounds [ratio]
    IF fDb >= 0.0 THEN
        FC_DL_AmpDbToRatio := DL_RATIO_MAX; // 按输入符号方向饱和至上限 [比] / saturate upward following the input sign [ratio]
    ELSE
        FC_DL_AmpDbToRatio := DL_RATIO_MIN; // 按输入符号方向饱和至下限 [比] / saturate downward following the input sign [ratio]
    END_IF
    eErr := 16#0001_01EC; // 溢出行为差异复用同一信息码，不另立码 / platform overflow difference reuses the same info id, no extra code
    bError := FALSE;      // 信息级不置故障 / info level never raises fault
    bValid := TRUE;       // 饱和值本身有效可用 / the saturated value itself is valid
    RETURN;               // 复检出口 / exit after the re-check
END_IF
eErr   := 0;     // 域内无错误 / in-domain, no error
bError := FALSE; // 信息级不置故障 / info level never raises fault
bValid := TRUE;  // 域内输出有效可用 / in-domain output is valid
END_FUNCTION

(* ---- FC_DL_AngleBisector.st ---- *)
(*==============================================================================
 * 名称 : FC_DL_AngleBisector —— 两角平分线（钝角取短弧中点，结果 [0,360)）
 * 分类 / 前缀 / 版本 : DL_MathData / FC_DL_ / 1.0.0
 * 溯源 : 开源语义参考（OSCAT/AixOCAT 族，MIT）或 clean-room IEC 实现，未复制源码
 * 平台 : 纯 IEC 61131-3
 * 功能说明 : 求 fA 与 fB 的角平分线：先取 fB-fA 的最短弧差 d∈[-180,180)
 *            （恒取短弧，即使两角相差为钝角侧也走短弧中点），平分角 =
 *            fA + 0.5*d，最后归一到 [0,360)。与 FC_DL_AngleLerpShort 的
 *            fT=0.5 特例一致，独立内联实现（无库内跨件依赖）。
 *            边界处理：任一输入非有限（NaN/±Inf）或 |角|>1.0E12 置 eErr 返回 0.0。
 * 错误码 : 16#0001_1B04 = 输入非有限（NaN/±Inf）或角度量超安全量程 ±1.0E12
 *          eErr=0 且 bValid=TRUE 表示返回值可用
 * 状态机 : R6 标注 N/A（纯函数无顺序状态，以本节替代 ELSE 兜底）
 * 红线 : R1/R2/R3 ✓ 零全局/零IO/纯IEC ｜ R4 ✓ 非有限拦截/量程防护 ｜ R10 ✓ 标准转换 ｜ R11 ✓ 分号收尾 ｜ R15 ✓ 无保留字撞名
 * 修订记录 : 2026-11-23 v1.0.0 首次入库（R76）
 *============================================================================*)
FUNCTION FC_DL_AngleBisector : LREAL
VAR_INPUT
    fA : LREAL;    // 角 A [度] / angle A in degrees
    fB : LREAL;    // 角 B [度] / angle B in degrees
END_VAR
VAR_OUTPUT
    eErr   : UDINT;    // 故障码，0=正常，1B04=输入非有限或超量程 / error code
    bError : BOOL;     // TRUE=本件发生故障 / TRUE when fault occurred
    bValid : BOOL;     // TRUE=返回值可用 / TRUE when return value is usable
END_VAR
VAR
    _d : LREAL;        // fB-fA 最短弧差 [度] / shortest-arc diff
    _m : LREAL;        // 平分角中间值 [度] / bisector raw value
END_VAR

FC_DL_AngleBisector := 0.0;                  // 返回值预设 0.0 / preset return to zero
eErr   := 16#0000_0000;                      // 故障码清零 / clear error code
bError := FALSE;                             // 故障标志清零 / clear error flag
bValid := TRUE;                              // 预设输出可用 / preset valid flag

IF (fA <> fA) OR ((fA - fA) <> (fA - fA))    // fA 非有限 / fA is NaN or infinite
   OR (fB <> fB) OR ((fB - fB) <> (fB - fB)) // fB 非有限 / fB is NaN or infinite
   OR (ABS(fA) > 1.0E12) OR (ABS(fB) > 1.0E12) THEN    // 角度量超安全量程 / beyond safe range
    eErr   := 16#0001_1B04;                  // 置故障码 / set error code
    bError := TRUE;                          // 置故障标志 / set error flag
    bValid := FALSE;                         // 返回值不可用 / return not usable
    RETURN;                                  // 返回 0.0 / return zero
END_IF

_d := fB - fA;                               // 原始差值 / raw difference
_d := _d - 360.0 * TRUNC(_d / 360.0);        // 整圈截断缩圈 / strip whole turns
IF _d >= 180.0 THEN                          // 上越界修正（恒取短弧）/ fix upper overflow
    _d := _d - 360.0;                        // 减一整圈 / subtract one turn
END_IF
IF _d < -180.0 THEN                          // 下越界修正 / fix lower overflow
    _d := _d + 360.0;                        // 加一整圈 / add one turn
END_IF

_m := fA + 0.5 * _d;                         // 短弧中点即平分角 / midpoint of short arc
_m := _m - 360.0 * TRUNC(_m / 360.0);        // 归一缩圈 / normalize by stripping turns
IF _m < 0.0 THEN                             // 负角修正 / fix negative angle
    _m := _m + 360.0;                        // 加一整圈 / add one turn
END_IF

FC_DL_AngleBisector := _m;                   // 回写 [0,360) 平分角 / write back bisector

END_FUNCTION

(* ---- FC_DL_AngleDiffRad.st ---- *)
(*
  ==================================================================
  组件名 Component  : FC_DL_AngleDiffRad
  分类   Category   : DL_MathData
  前缀   Naming     : FC_DL_ ｜ b/n/u/f 类型前缀制（R265）
  版本   Version    : 1.0.0
  功能   Purpose    : 两弧度角最短带符号差：fDiff = fAngleA − fAngleB 归一
                      至 [−π, π]。回绕处理两步：先 TRUNC 整圈数把差值压入
                      (−2π, 2π)（TRUNC 向零取整，余数保号），再按 ±π 边界
                      单次平移进 [−π, π]。跨 ±π 回绕（359°→1° 类）输出 ≈
                      −0.035 而非 ≈ 6.26。超大量级角（|差| > π·2^52）精
                      度受 LREAL 整数位尾差限制，头注声明为固有边界。
  来源   Source     : t2-1-lgf-math（角度最短差归一为公开数学口径
                      （mod-2π 最短代表元），实现零源码复制）
  互引   Cross-ref  : FC_DL_AngleDiffWrap / FC_DL_WrapAngleDeg（既有角度
                      族邻件：Wrap 件为角度自身回绕，本件为两角差值归一，
                      弧度口径属主；度口径见 WrapAngleDeg）
  平台   Platform   : 纯 IEC 61131-3 四则 + ABS/TRUNC，三平台通用
  依赖   Depends    : 无 DL_ 内部依赖；无标准库
  红线   Redline    : R1 零全局/VAR_EXTERNAL/R2 零 %I/%Q/R3 纯 IEC 标准
                      R4 非有限闸 + 输出域显式（[−π,π] 复核）/R5 全变量
                      双语同行注释/R6 纯函数无状态机（CASE 不适用）
                      /R7 无定时器与沿检测/R8 阈值全常量化
  错误码 Codes      : 01【失效级】任一输入角非有限（NaN 自反判 / Inf 上限
                      兜底判），返回 0
                      02【失效级】归一后输出越出 [−π−ε, π+ε] 域（结构性
                      罕见兜底），返回 0
  码位反证 Note     : 01/02 分立依据（R90）：01 在输入面、02 在输出域面
                      可观测；02 若并入 01，则「回绕算法自身失效」这一信
                      号将不可观测，故必须分立。
  验收   Acceptance : V1 A=0.1,B=−0.1 → 0.2 ｜ V2 A=6.26,B=0.02 → ≈−0.04
                      （跨 π 回绕）｜ V3 A=−3.2,B=3.2 → ≈3.083（跨 −π）
                      ｜ V4 A=B+2π → ≈0 ｜ V5 含 NaN → 码 01
  变更   Revision   : 2026-11-22  v1.0.0  R67 首版（编码阶段批 2 序 2）
  ==================================================================
*)
FUNCTION FC_DL_AngleDiffRad : LREAL
VAR_INPUT
    fAngleA : LREAL;  // 角 A [rad] / the angle A in radians
    fAngleB : LREAL;  // 角 B [rad] / the angle B in radians
END_VAR
VAR_OUTPUT
    bValid  : BOOL;   // 差值可用标志 [-] / the difference usable flag
    nErrId  : UDINT;  // 错误码，0=正常，01/02 见头注 [码] / the error code [code]
END_VAR
VAR
    fD      : LREAL;  // 原始差值工作寄存器 [rad] / the raw difference register
    nTurn   : LREAL;  // 整圈数工作寄存器（TRUNC 向零取整）/ the full turn count register
END_VAR
VAR CONSTANT
    ADR_PI       : LREAL := 3.141592653589793;     // π [rad] / the pi constant
    ADR_TWO_PI   : LREAL := 6.283185307179586;     // 2π [rad] / the two pi constant
    ADR_EPS      : LREAL := 1.0E-9;                // 输出域复核容差 [rad] / the output domain tolerance
    ADR_FIN_MAX  : LREAL := 1.7976931348623157E308; // LREAL 有限上限 / the finite LREAL limit
    ADR_ERR_NONE : UDINT := 16#0000_0000;          // 无错误 [码] / no error [code]
    ADR_ERR_NAN  : UDINT := 16#0000_0001;          // 码 01：输入非有限 / code 01, non finite input
    ADR_ERR_DOM  : UDINT := 16#0000_0002;          // 码 02：输出域越界 / code 02, output domain breach
END_VAR

// 段 1｜输出预置 / segment 1, preset the outputs
FC_DL_AngleDiffRad := 0.0;  // 失效缺省返回 0 / fault default returns zero
bValid := FALSE;            // 预置不可用 / preset unusable
nErrId := ADR_ERR_NONE;     // 预置无错误 / preset no error

// 段 2｜输入非有限闸（码 01）/ segment 2, the input finite gate
IF (fAngleA <> fAngleA) OR (fAngleB <> fAngleB)
   OR (ABS(fAngleA) > ADR_FIN_MAX) OR (ABS(fAngleB) > ADR_FIN_MAX) THEN
    nErrId := ADR_ERR_NAN;
    RETURN;
END_IF

// 段 3｜原始差值与整圈归约（TRUNC 向零取整，余数保号压入 (−2π, 2π)）
//      segment 3, the raw difference and the full turn reduction
fD := fAngleA - fAngleB;                  // 原始差 [rad] / the raw difference
nTurn := TRUNC(fD / ADR_TWO_PI);          // 整圈数（LREAL 口径，不进 DINT 溢出面）/ the turn count
fD := fD - nTurn * ADR_TWO_PI;            // 压入 (−2π, 2π) / reduce into the open two pi band

// 段 4｜半圈平移进 [−π, π]（单次判界，无循环）/ segment 4, the half turn shift into the pi band
IF fD > ADR_PI THEN                       // 正侧越界回绕 / the positive wrap
    fD := fD - ADR_TWO_PI;
ELSIF fD < -ADR_PI THEN                  // 负侧越界回绕 / the negative wrap
    fD := fD + ADR_TWO_PI;
END_IF

// 段 5｜输出域复核（码 02）与出口 / segment 5, the output domain recheck and exit
IF (fD <> fD) OR (fD < -ADR_PI - ADR_EPS) OR (fD > ADR_PI + ADR_EPS) THEN
    nErrId := ADR_ERR_DOM;                // 归一后仍越域（结构性罕见兜底）/ the breach after reduction
    RETURN;
END_IF
FC_DL_AngleDiffRad := fD;                 // 最短带符号差 [rad] / the shortest signed difference
bValid := TRUE;                           // 差值可用 / the difference is usable
END_FUNCTION

(* ---- FC_DL_AngleDiffWrap.st ---- *)
(*
  FC_DL_AngleDiffWrap  —  角度差环绕归一至 ±180° / Angle difference wrapped into the plus-minus 180 degree span
  分类 Category : DL_MathData
  版本 Version  : 1.0.0
  来源 Source   : iec-std-wrapper — 标准语义包装族（fMod 归一口径），IEC 61131-3 标准语义的道莅防御性实现
  溯源 Origin   : clean-room 实现，未复制任何源码行
  功能 Function : 1) 返回 fAngA - fAngB 归一至 [-180.0, 180.0] 的环绕角差 [deg]；
                  2) 归一口径：先 fMod := 差值 - 360 × TRUNC(差值/360)（fMod 语义），
                  再 fMod > 180 减 360、fMod <= -180 加 360，360° 环绕；
                  3) 进位点向量：正好 ±180.0（含 -180 精确落点）一律归 +180.0，不归 -180.0；
                  4) 非有限输入（NaN 自反判 / Inf 差值自减判）→ 返回 0、故障级 03E0、bValid FALSE。
  边界 Boundary : ① 非有限判定：NaN 用 x <> x 自反判；Inf 用 (x-x) <> (x-x) 判，
                  禁近似阈值（R40 LREAL 口径）；
                  ② 浮点比较禁用 = / <> 判相等（除自反 NaN 判外），进位点用容差 1.0E-6；
                  ③ 无 GVL 依赖：纯函数，无外部变量引用，无物理 IO 地址；
                  ④ 返回角差量纲 [deg]，输入量纲亦须 [deg]，换算由调用方完成。
  依赖 Depends  : 仅 Standard.library（TRUNC / ABS / LREAL 算术）
  码表 Error codes（段 0001，窗口 03E0 / 04A3）:
    16#0001_03E0 故障级：输入非有限（NaN 或 Inf），返回 0，bValid = FALSE，bError = TRUE
    16#0001_04A3 信息级：进位点命中（|结果| = 180.0 容差内，归 +180）
  修订历史 Revision :
    2026-11-19  v1.0.0  R41 首版（批次 1 · 序号 3；同日机检后主控重建正文，规格以本头注释为准）
*)

FUNCTION FC_DL_AngleDiffWrap : LREAL
VAR_INPUT
    fAngA       : LREAL;             // 角 A [deg]，量纲须为度 / Angle A in degrees
    fAngB       : LREAL;             // 角 B [deg]，量纲须为度 / Angle B in degrees
END_VAR
VAR_OUTPUT
    eErr        : UDINT;             // 事件码，0 = 正常 / Event code
    bError      : BOOL;              // 故障级标志 / Fault-level flag
    bValid      : BOOL;              // 返回值是否可用 / Result usable flag
END_VAR
VAR
    fDiff       : LREAL;             // 原始差值 [deg] / Raw difference before wrap
    fMod        : LREAL;             // 模 360 中间量 [deg] / Modulo-360 intermediate
END_VAR
VAR CONSTANT
    DL_ADW_TOL       : LREAL := 1.0E-6;         // 进位点容差 [deg] / Tie-point tolerance
    DL_ADW_ERR_NFIN  : UDINT := 16#0001_03E0;   // 故障级：输入非有限 / Fault: non-finite input
    DL_ADW_INFO_TIE  : UDINT := 16#0001_04A3;   // 信息级：进位点命中 / Info: tie-point hit
END_VAR

(* —— 段 1｜返回值与错误状态预置 —— *)
FC_DL_AngleDiffWrap := 0.0;         // 缺省返回 0 / default return zero
eErr := 16#0000_0000;               // 预置无事件 / preset no event
bError := FALSE;                    // 预置无故障 / preset no fault
bValid := FALSE;                    // 预置不可用 / preset unusable

(* —— 段 2｜非有限输入拦截（NaN 自反判 / Inf 差值自减判，R40 LREAL 口径）—— *)
IF (fAngA <> fAngA) OR (fAngB <> fAngB)
   OR ((fAngA - fAngA) <> (fAngA - fAngA))
   OR ((fAngB - fAngB) <> (fAngB - fAngB)) THEN
    FC_DL_AngleDiffWrap := 0.0;     // 非有限输入返回 0 / non-finite input returns zero
    eErr := DL_ADW_ERR_NFIN;        // 置故障级 03E0 / fault code 03E0
    bError := TRUE;                 // 故障标志 / fault flag
    bValid := FALSE;                // 结果不可用 / result unusable
    RETURN;
END_IF

(* —— 段 3｜域内归一（委托 fMod 语义：TRUNC 取整方向与 fMod 一致）—— *)
fDiff := fAngA - fAngB;             // 原始差值 / raw difference
fMod := fDiff - 360.0 * TRUNC(fDiff / 360.0);   // fMod 语义归一 / fMod-semantics normalize
IF fMod > 180.0 THEN                // (180, 360) 区间减一圈 / wrap upper half
    fMod := fMod - 360.0;
END_IF
IF fMod <= -180.0 THEN              // [-360, -180] 区间加一圈（-180 精确落点归 +180）/ wrap lower half
    fMod := fMod + 360.0;
END_IF

(* —— 段 4｜进位点向量：±180 精确落点一律归 +180.0 —— *)
IF ABS(ABS(fMod) - 180.0) <= DL_ADW_TOL THEN    // 容差内视为进位点 / within tolerance is tie point
    fMod := 180.0;                  // 统一归 +180 / unify to +180
    eErr := DL_ADW_INFO_TIE;        // 置信息级 04A3 / info code 04A3
END_IF

(* —— 段 5｜结果复检兜底（防溢出/异常传播）—— *)
IF (fMod <> fMod) OR (fMod < -180.0) OR (fMod > 180.0) THEN
    FC_DL_AngleDiffWrap := 0.0;     // 复检失败返回 0 / recheck failed returns zero
    eErr := DL_ADW_ERR_NFIN;        // 归故障级 / fault-level
    bError := TRUE;
    bValid := FALSE;
    RETURN;
END_IF

FC_DL_AngleDiffWrap := fMod;        // 输出环绕角差 / output wrapped difference
bError := FALSE;                    // 无故障 / no fault
bValid := TRUE;                     // 结果可用 / result usable

END_FUNCTION
